(* IEC 61131-3 sources: plc_NativeGateway/src (part 2) *)

(* ---- NG_HmiEdit.st ---- *)
FUNCTION_BLOCK NG_HmiEdit
VAR_INPUT
    Busy : BOOL;
    StoreBusy : BOOL;
    Managed : BOOL;
    LocalRevision : ULINT;
    NowMs : ULINT;
END_VAR
VAR_IN_OUT
    Hmi : NG_Hmi;
    Active : NG_Config;
    Bootstrap : NG_Bootstrap;
    States : ARRAY[1..50] OF NG_MeterState;
    Samples : ARRAY[1..320] OF NG_Sample;
END_VAR
VAR_OUTPUT
    Submit : BOOL;
    SubmitBroker : BOOL;
    SubmitMode : BOOL;
    SubmitReset : BOOL;
    ClearConfig : BOOL;
    Draft : NG_Config;
    NewBroker : NG_Bootstrap;
    NewManaged : BOOL;
END_VAR
VAR
    Change : NG_EditDevice;
    EditPoints : ARRAY[1..32] OF NG_Point;
    BlankPoint : NG_Point;
    BlankDevice : NG_Device;
    BaseVersion : ULINT;
    BaseRevision : ULINT;
    ModeTargetManaged : BOOL;
    ModeReviewOpen : BOOL;
    ResetReviewOpen : BOOL;
    Initialized : BOOL;
    Dirty : BOOL;
    Awaiting : BOOL;
    Reload : BOOL;
    LoadDevice : BOOL;
    LoadPoint : BOOL;
    ValidBroker : BOOL;
    RefreshAt : ULINT;
    Nav : STRING[16];
    d : INT;
    p : INT;
    i : INT;
    row : INT;
    a : INT;
    b : INT;
    idx : INT;
    pages : INT;
    point : NG_Point;
    device : NG_Device;
    rows : ARRAY[1..8] OF NG_UiLabel;
    marker : STRING[3];
    status : STRING[24];
    value : STRING[64];
    cmd : BOOL;
    Utf8 : NG_Utf8Label;
    DeviceLabel : NG_UiLabel;
    PointLabel : NG_UiLabel;
    UnitLabel : NG_UiLabel;
END_VAR
Submit := FALSE; SubmitBroker := FALSE; SubmitMode := FALSE; SubmitReset := FALSE; ClearConfig := FALSE; LoadDevice := FALSE; LoadPoint := FALSE;
Nav := Hmi.Navigation; Hmi.Navigation := '';
IF Nav='ZH' THEN Hmi.English:=FALSE;
ELSIF Nav='EN' THEN Hmi.English:=TRUE;
ELSIF Nav='REFRESH' THEN IF Dirty THEN Hmi.View:=5; ELSE Hmi.Load:=TRUE; END_IF;
ELSIF Nav='DISCARD' THEN Hmi.Load:=TRUE; Hmi.View:=0;
ELSIF Nav='REVIEW' THEN Hmi.View:=6;
ELSIF Nav='COMMIT' THEN Hmi.Apply:=TRUE;
ELSIF Nav='DEVON' THEN Hmi.DeviceEnabled:='true';
ELSIF Nav='DEVOFF' THEN Hmi.DeviceEnabled:='false';
ELSIF Nav='POINTON' THEN Hmi.PointEnabled:='true';
ELSIF Nav='POINTOFF' THEN Hmi.PointEnabled:='false';
ELSIF Nav='MODEPAGE' THEN ModeReviewOpen:=FALSE; ResetReviewOpen:=FALSE; Hmi.View:=13;
ELSIF Nav='MODEHUB' THEN ModeTargetManaged:=TRUE; ModeReviewOpen:=TRUE; ResetReviewOpen:=FALSE; Hmi.ClearOnMaintenance:=FALSE; Hmi.View:=15;
ELSIF Nav='MODELOCAL' THEN ModeTargetManaged:=FALSE; ModeReviewOpen:=TRUE; ResetReviewOpen:=FALSE; Hmi.ClearOnMaintenance:=FALSE; Hmi.View:=14;
ELSIF Nav='MODEKEEP' THEN Hmi.ClearOnMaintenance:=FALSE;
ELSIF Nav='MODECLEAR' THEN Hmi.ClearOnMaintenance:=TRUE;
ELSIF Nav='MODECOMMIT' THEN
    IF ModeReviewOpen AND ((Hmi.View=14) OR (Hmi.View=15)) THEN Hmi.SwitchMode:=TRUE;
    ELSE Hmi.Status:='Open the management mode confirmation before saving.'; END_IF;
ELSIF Nav='RESETPAGE' THEN ModeReviewOpen:=FALSE; ResetReviewOpen:=TRUE; Hmi.View:=16;
ELSIF Nav='RESETCOMMIT' THEN
    IF ResetReviewOpen AND (Hmi.View=16) THEN
        IF StoreBusy THEN Hmi.Status:='Busy: configuration transaction in progress. Try again shortly.';
        ELSE SubmitReset:=TRUE; ResetReviewOpen:=FALSE; Dirty:=FALSE; Awaiting:=FALSE; Reload:=TRUE; Hmi.View:=0; Hmi.Status:='Clearing local configuration and version baseline...'; END_IF;
    ELSE Hmi.Status:='Open the reset confirmation before clearing local configuration.'; END_IF;
ELSIF Nav='CYCLIC' THEN Hmi.ReportMode:='cyclic';
ELSIF Nav='CHANGE' THEN Hmi.ReportMode:='change';
ELSIF Nav='BOTH' THEN Hmi.ReportMode:='change_or_cyclic';
ELSIF Nav='HOLDING' THEN Hmi.Area:='holding_register';
ELSIF Nav='INPUT' THEN Hmi.Area:='input_register';
ELSIF Nav='COIL' THEN Hmi.Area:='coil';
ELSIF Nav='DISCRETE' THEN Hmi.Area:='discrete_input';
ELSIF Nav='UINT16' THEN Hmi.DataType:='uint16'; Hmi.ByteOrder:='AB';
ELSIF Nav='INT16' THEN Hmi.DataType:='int16'; Hmi.ByteOrder:='AB';
ELSIF Nav='UINT32' THEN Hmi.DataType:='uint32'; Hmi.ByteOrder:='ABCD';
ELSIF Nav='INT32' THEN Hmi.DataType:='int32'; Hmi.ByteOrder:='ABCD';
ELSIF Nav='FLOAT32' THEN Hmi.DataType:='float32'; Hmi.ByteOrder:='ABCD';
ELSIF Nav='BOOL' THEN Hmi.DataType:='bool'; Hmi.ByteOrder:=''; Hmi.Scale:='1'; Hmi.Offset:='0'; Hmi.Deadband:='0';
ELSIF Nav='ADVANCED' THEN Hmi.Advanced:=NOT Hmi.Advanced;
ELSIF Nav='BROKERREVIEW' THEN Hmi.View:=7;
ELSIF Nav='BROKERCOMMIT' THEN Hmi.SaveBroker:=TRUE;
ELSIF Nav='HELP' THEN Hmi.View:=8;
ELSIF Nav='TYPEPICK' THEN Hmi.View:=9;
ELSIF Nav='AREAPICK' THEN Hmi.View:=10;
ELSIF Nav='REPORTPICK' THEN Hmi.View:=11;
ELSIF Nav='GATEWAY' THEN Hmi.View:=12;
ELSIF Nav='POINTBACK' THEN Hmi.View:=2;
END_IF;
IF (Nav='CYCLIC') OR (Nav='CHANGE') OR (Nav='BOTH') OR (Nav='HOLDING') OR (Nav='INPUT') OR (Nav='COIL') OR (Nav='DISCRETE') OR (Nav='UINT16') OR (Nav='INT16') OR (Nav='UINT32') OR (Nav='INT32') OR (Nav='FLOAT32') OR (Nav='BOOL') THEN Hmi.View:=2; END_IF;
Hmi.Managed:=Managed;
IF Managed THEN Hmi.ManagementMode:='HUB_MANAGED'; ELSE Hmi.ManagementMode:='STANDALONE'; END_IF;
IF Managed AND ((Nav='DNEW') OR (Nav='PNEW') OR (Nav='DDEL') OR (Nav='PDEL') OR (Nav='PERIOD') OR Hmi.SaveDevice OR Hmi.SavePoint OR Hmi.RemoveDevice OR Hmi.RemovePoint OR Hmi.Apply) THEN
    Nav := ''; Hmi.SaveDevice:=FALSE; Hmi.SavePoint:=FALSE; Hmi.RemoveDevice:=FALSE; Hmi.RemovePoint:=FALSE; Hmi.Apply:=FALSE;
    Hmi.View:=0; Hmi.Status:='HUB_MANAGED: publish device and point changes from Hub.';
END_IF;
IF Managed THEN Hmi.ConfigSource:='HUB_MANAGED - local device/point changes blocked'; ELSE Hmi.ConfigSource:='MAINTENANCE - incoming platform configuration locked'; END_IF;
IF NOT Initialized THEN Reload := TRUE; Initialized := TRUE; END_IF;
IF Awaiting AND (Active.Version = Draft.Version) AND NOT Busy THEN Dirty := FALSE; Awaiting := FALSE; Reload := TRUE; Hmi.View:=0; END_IF;
IF ((Active.Version <> BaseVersion) OR (LocalRevision <> BaseRevision)) AND NOT Dirty AND NOT Awaiting AND NOT Busy THEN Reload := TRUE; END_IF;
IF Hmi.Load AND NOT Busy THEN Reload := TRUE; Hmi.View:=0; Hmi.Status := 'Display refreshed from active configuration. Unapplied draft discarded.'; END_IF;
IF Reload THEN
    Draft := Active; BaseVersion := Active.Version; BaseRevision := LocalRevision; Dirty := FALSE; Reload := FALSE;
    Hmi.Enabled := TO_STRING(Draft.enabled,''); Hmi.BatchIntervalMs := TO_STRING(Draft.batchIntervalMs,'{0:d}'); Hmi.MaxBatchPoints := TO_STRING(Draft.maxBatchPoints,'{0:d}');
    IF NOT NG_Range(Hmi.DeviceIndex,1,50,TRUE) THEN Hmi.DeviceIndex := '1'; END_IF;
    Hmi.PointIndex := '1'; LoadDevice := TRUE; LoadPoint := TRUE;
END_IF;
d := 1; p := 1;
IF NG_Range(Hmi.DeviceIndex,1,50,TRUE) THEN d := TO_INT(Hmi.DeviceIndex); END_IF;
IF NG_Range(Hmi.PointIndex,1,32,TRUE) THEN p := TO_INT(Hmi.PointIndex); END_IF;
IF Nav = 'LIST' THEN Hmi.View := 0;
ELSIF Nav = 'MQTT' THEN Hmi.View := 3;
ELSIF Nav = 'DEDIT' THEN Hmi.View := 1; LoadDevice := TRUE;
ELSIF Nav = 'PEDIT' THEN Hmi.View := 2; LoadPoint := TRUE;
ELSIF Nav = 'DPREV' THEN Hmi.DevicePage := MAX(1,Hmi.DevicePage-1);
ELSIF Nav = 'DNEXT' THEN Hmi.DevicePage := MIN(MAX(1,(Draft.DeviceCount+7)/8),Hmi.DevicePage+1);
ELSIF Nav = 'PPREV' THEN Hmi.PointPage := MAX(1,Hmi.PointPage-1);
ELSIF Nav = 'PNEXT' THEN IF d <= Draft.DeviceCount THEN Hmi.PointPage := MIN(MAX(1,(Draft.Devices[d].PointCount+7)/8),Hmi.PointPage+1); END_IF;
ELSIF Nav = 'DDEL' THEN Hmi.DeleteKind := 1; Hmi.View := 4;
ELSIF Nav = 'PDEL' THEN Hmi.DeleteKind := 2; Hmi.View := 4;
ELSIF Nav = 'CANCEL' THEN Hmi.DeleteKind := 0; Hmi.View := 0;
ELSIF Nav = 'DNEW' THEN
    IF Draft.DeviceCount >= 50 THEN Hmi.Status := 'Capacity reached: 50 devices.';
    ELSE
        d := Draft.DeviceCount+1; Hmi.DeviceIndex := TO_STRING(d,'{0:d}'); Hmi.PointIndex := '1'; Hmi.View := 1;
        Hmi.DeviceId := CONCAT('meter-',TO_STRING(d,'{0:d}')); Hmi.DeviceName := CONCAT('Meter ',TO_STRING(d,'{0:d}'));
        Hmi.Host := '192.168.0.5'; Hmi.Port := '11502'; Hmi.UnitId := TO_STRING(d,'{0:d}'); Hmi.DeviceEnabled := 'true';
        Hmi.ConnectTimeoutMs := '3000'; Hmi.RequestTimeoutMs := '1500'; Hmi.RetryCount := '0';
        Hmi.Status := 'New device: save into draft, then add its points.';
    END_IF;
ELSIF Nav = 'PNEW' THEN
    IF d > Draft.DeviceCount THEN Hmi.Status := 'Save a device into the draft first.';
    ELSIF (Draft.Devices[d].PointCount >= 32) OR (Draft.PointCount >= 320) THEN Hmi.Status := 'Capacity reached: 32 points/device, 320 shared points.';
    ELSE
        p := Draft.Devices[d].PointCount+1; Hmi.PointIndex := TO_STRING(p,'{0:d}'); Hmi.View := 2;
        Hmi.PointId := CONCAT('point-',TO_STRING(p,'{0:d}')); Hmi.PointName := CONCAT('Point ',TO_STRING(p,'{0:d}')); Hmi.PointEnabled := 'true';
        Hmi.DataType := 'float32'; Hmi.Area := 'input_register'; Hmi.Address := TO_STRING((p-1)*2,'{0:d}'); Hmi.ByteOrder := 'ABCD';
        Hmi.PollIntervalMs := '5000'; Hmi.ReportIntervalMs := '5000'; Hmi.Scale := '1'; Hmi.Offset := '0'; Hmi.Unit := '';
        Hmi.ReportMode := 'cyclic'; Hmi.Deadband := '0'; Hmi.StaleAfterMs := '20000';
        Hmi.Status := 'New point: save into draft, then apply the complete draft.';
    END_IF;
ELSIF LEN(Nav) = 2 THEN
    IF (LEFT(Nav,1) = 'D') AND NG_Range(RIGHT(Nav,1),1,8,TRUE) THEN
        i := (Hmi.DevicePage-1)*8+TO_INT(RIGHT(Nav,1));
        IF i <= Draft.DeviceCount THEN d := i; p := 1; Hmi.DeviceIndex := TO_STRING(d,'{0:d}'); Hmi.PointIndex := '1'; Hmi.PointPage := 1; LoadDevice := TRUE; LoadPoint := TRUE; END_IF;
    ELSIF (LEFT(Nav,1) = 'P') AND NG_Range(RIGHT(Nav,1),1,8,TRUE) AND (d <= Draft.DeviceCount) THEN
        i := (Hmi.PointPage-1)*8+TO_INT(RIGHT(Nav,1));
        IF i <= Draft.Devices[d].PointCount THEN p := i; Hmi.PointIndex := TO_STRING(p,'{0:d}'); LoadPoint := TRUE; END_IF;
    END_IF;
END_IF;
IF LoadDevice AND (d <= Draft.DeviceCount) THEN
    device := Draft.Devices[d];
    Hmi.DeviceId := device.deviceId; Hmi.DeviceName := device.name; Hmi.DeviceEnabled := TO_STRING(device.enabled,''); Hmi.Host := device.host;
    Hmi.Port := TO_STRING(device.port,'{0:d}'); Hmi.UnitId := TO_STRING(device.unitId,'{0:d}'); Hmi.ConnectTimeoutMs := TO_STRING(device.connectTimeoutMs,'{0:d}');
    Hmi.RequestTimeoutMs := TO_STRING(device.requestTimeoutMs,'{0:d}'); Hmi.RetryCount := TO_STRING(device.retryCount,'{0:d}');
END_IF;
IF Hmi.LoadPoint THEN LoadPoint := TRUE; END_IF;
IF LoadPoint AND (d <= Draft.DeviceCount) THEN
    IF p <= Draft.Devices[d].PointCount THEN
        point := Draft.Points[Draft.Devices[d].PointStart+p-1];
        Hmi.PointId := point.pointId; Hmi.PointName := point.name; Hmi.PointEnabled := TO_STRING(point.enabled,''); Hmi.DataType := point.dataType;
        Hmi.PollIntervalMs := TO_STRING(point.pollIntervalMs,'{0:d}'); Hmi.ReportIntervalMs := TO_STRING(point.reportIntervalMs,'{0:d}');
        Hmi.Scale := TO_STRING(point.scale,'{0:F6}'); Hmi.Offset := TO_STRING(point.offset,'{0:F6}'); Hmi.Unit := point.unit; Hmi.ReportMode := point.reportMode;
        Hmi.Deadband := TO_STRING(point.deadband,'{0:F6}'); Hmi.StaleAfterMs := TO_STRING(point.staleAfterMs,'{0:d}'); Hmi.Area := point.area;
        Hmi.Address := TO_STRING(point.address,'{0:d}'); Hmi.ByteOrder := point.byteOrder;
        Hmi.DevicePollMs := Hmi.PollIntervalMs; Hmi.DeviceReportMs := Hmi.ReportIntervalMs;
    END_IF;
END_IF;
cmd := Hmi.SaveDevice OR Hmi.SavePoint OR Hmi.RemoveDevice OR Hmi.RemovePoint OR Hmi.Apply OR Hmi.SaveBroker OR Hmi.SwitchMode OR (Nav = 'PERIOD');
IF cmd AND ((Hmi.SaveBroker AND StoreBusy) OR ((NOT Hmi.SaveBroker) AND Busy)) THEN Hmi.Status := 'Busy: configuration transaction in progress. Try again shortly.';
ELSIF cmd THEN
    IF NOT NG_Range(Hmi.DeviceIndex,1,50,TRUE) OR NOT NG_Range(Hmi.PointIndex,1,32,TRUE) THEN Hmi.Status := 'Device index 1..50; point index 1..32.';
    ELSE
        d := TO_INT(Hmi.DeviceIndex); p := TO_INT(Hmi.PointIndex); device := BlankDevice;
        IF d <= Draft.DeviceCount THEN device := Draft.Devices[d]; FOR i := 1 TO device.PointCount DO EditPoints[i] := Draft.Points[device.PointStart+i-1]; END_FOR; END_IF;
        IF Hmi.SaveDevice THEN
            IF (d > Draft.DeviceCount+1) OR NOT NG_ValidId(Hmi.DeviceId) OR (LEN(Hmi.DeviceName)=0) OR NOT NG_IPv4(Hmi.Host) OR
               NOT NG_Range(Hmi.Port,1,65535,TRUE) OR NOT NG_Range(Hmi.UnitId,0,255,TRUE) OR NOT NG_Range(Hmi.ConnectTimeoutMs,1,300000,TRUE) OR NOT NG_Range(Hmi.RequestTimeoutMs,1,300000,TRUE) OR NOT NG_Range(Hmi.RetryCount,0,10,TRUE) THEN Hmi.Status := 'Invalid device fields: check ID, name, IPv4, port and timeout values.';
            ELSE
                device.deviceId := Hmi.DeviceId; device.name := Hmi.DeviceName; device.enabled := (Hmi.DeviceEnabled='true') OR (Hmi.DeviceEnabled='TRUE');
                device.host := Hmi.Host; device.port := TO_UINT(Hmi.Port); device.unitId := TO_USINT(Hmi.UnitId); device.connectTimeoutMs := TO_UDINT(Hmi.ConnectTimeoutMs);
                device.requestTimeoutMs := TO_UDINT(Hmi.RequestTimeoutMs); device.retryCount := TO_USINT(Hmi.RetryCount);
                Change(DeviceIndex := d, Remove := FALSE, Replacement := device, Config := Draft, Points := EditPoints);
                IF Change.ErrorText = '' THEN Dirty := TRUE; Hmi.View := 0; Hmi.Status := 'Device saved to draft. Apply draft to persist.'; ELSE Hmi.Status := Change.ErrorText; END_IF;
            END_IF;
        END_IF;
        IF Hmi.SavePoint THEN
            IF (d > Draft.DeviceCount) OR (p > device.PointCount+1) OR NOT NG_ValidId(Hmi.PointId) OR (LEN(Hmi.PointName)=0) OR
               NOT NG_Range(Hmi.PollIntervalMs,1,86400000,TRUE) OR NOT NG_Range(Hmi.ReportIntervalMs,1,86400000,TRUE) OR NOT NG_Range(Hmi.StaleAfterMs,1,86400000,TRUE) OR NOT NG_Range(Hmi.Address,0,65535,TRUE) OR
               NOT NG_Range(Hmi.Scale,-1.0E20,1.0E20,FALSE) OR NOT NG_Range(Hmi.Offset,-1.0E20,1.0E20,FALSE) OR NOT NG_Range(Hmi.Deadband,0,1.0E20,FALSE) THEN Hmi.Status := 'Invalid point fields; save the device first and check numeric fields.';
            ELSE
                point := BlankPoint; point.pointId := Hmi.PointId; point.name := Hmi.PointName; point.enabled := (Hmi.PointEnabled='true') OR (Hmi.PointEnabled='TRUE');
                point.dataType := Hmi.DataType; point.pollIntervalMs := TO_UDINT(Hmi.PollIntervalMs); point.reportIntervalMs := TO_UDINT(Hmi.ReportIntervalMs);
                point.scale := TO_LREAL(Hmi.Scale); point.offset := TO_LREAL(Hmi.Offset); point.unit := Hmi.Unit; point.reportMode := Hmi.ReportMode;
                point.deadband := TO_LREAL(Hmi.Deadband); point.staleAfterMs := TO_UDINT(Hmi.StaleAfterMs); point.area := Hmi.Area; point.address := TO_UINT(Hmi.Address); point.byteOrder := Hmi.ByteOrder;
                EditPoints[p] := point; IF p > device.PointCount THEN device.PointCount := p; END_IF;
                Change(DeviceIndex := d, Remove := FALSE, Replacement := device, Config := Draft, Points := EditPoints);
                IF Change.ErrorText = '' THEN Dirty := TRUE; Hmi.View := 0; Hmi.Status := 'Point saved to draft. Apply draft to persist.'; ELSE Hmi.Status := Change.ErrorText; END_IF;
            END_IF;
        END_IF;
        IF Hmi.RemoveDevice AND (d <= Draft.DeviceCount) THEN
            Change(DeviceIndex := d, Remove := TRUE, Replacement := device, Config := Draft, Points := EditPoints);
            IF Change.ErrorText = '' THEN Dirty := TRUE; Hmi.DeviceIndex := '1'; Hmi.PointIndex := '1'; Hmi.View := 0; Hmi.DeleteKind := 0; Hmi.Status := 'Device and points removed from draft. Apply to persist.'; END_IF;
        END_IF;
        IF Hmi.RemovePoint AND (d <= Draft.DeviceCount) AND (p <= device.PointCount) THEN
            FOR i := p TO device.PointCount-1 DO EditPoints[i] := EditPoints[i+1]; END_FOR; device.PointCount := device.PointCount-1;
            Change(DeviceIndex := d, Remove := FALSE, Replacement := device, Config := Draft, Points := EditPoints);
            IF Change.ErrorText = '' THEN Dirty := TRUE; Hmi.PointIndex := '1'; Hmi.View := 0; Hmi.DeleteKind := 0; Hmi.Status := 'Point removed from draft. Apply to persist.'; END_IF;
        END_IF;
        IF (Nav = 'PERIOD') AND (d <= Draft.DeviceCount) THEN
            IF NOT NG_Range(Hmi.DevicePollMs,1,28800000,TRUE) OR NOT NG_Range(Hmi.DeviceReportMs,1,86400000,TRUE) THEN Hmi.Status := 'Invalid device polling/report period.';
            ELSE
                FOR i := 1 TO device.PointCount DO idx := device.PointStart+i-1; Draft.Points[idx].pollIntervalMs := TO_UDINT(Hmi.DevicePollMs); Draft.Points[idx].reportIntervalMs := TO_UDINT(Hmi.DeviceReportMs); Draft.Points[idx].staleAfterMs := MAX(Draft.Points[idx].staleAfterMs,Draft.Points[idx].pollIntervalMs*3); END_FOR;
                Dirty := TRUE; Hmi.Status := 'Device point periods updated in draft. Apply to persist.';
            END_IF;
        END_IF;
        IF Hmi.Apply THEN
            IF (BaseVersion <> Active.Version) OR (BaseRevision <> LocalRevision) THEN Hmi.Status := 'VERSION_CONFLICT: reload active configuration before applying.';
            ELSIF NOT NG_Range(Hmi.BatchIntervalMs,1,86400000,TRUE) OR NOT NG_Range(Hmi.MaxBatchPoints,1,64,TRUE) THEN Hmi.Status := 'Invalid gateway batch settings.';
            ELSE
                Draft.enabled := (Hmi.Enabled='true') OR (Hmi.Enabled='TRUE'); Draft.batchIntervalMs := TO_UDINT(Hmi.BatchIntervalMs); Draft.maxBatchPoints := TO_UINT(Hmi.MaxBatchPoints); Hmi.Status := NG_CheckConfig(Draft);
                IF Hmi.Status = '' THEN Draft.Version := Active.Version; Submit := TRUE; Awaiting := TRUE; Dirty := TRUE; Hmi.Status := 'Saving, hashing and reading back configuration...'; END_IF;
            END_IF;
        END_IF;
        IF Hmi.SwitchMode THEN
            NewManaged := ModeTargetManaged;
            IF NewManaged = Managed THEN Hmi.Status := 'The selected management mode is already active.';
            ELSE
                ClearConfig := NOT NewManaged AND Hmi.ClearOnMaintenance;
                SubmitMode := TRUE; ModeReviewOpen:=FALSE; Dirty := FALSE; Awaiting := FALSE; Reload := TRUE;
                Hmi.View := 13; Hmi.Status := 'Saving management mode; existing identity is retained.';
            END_IF;
        END_IF;
        IF Hmi.SaveBroker THEN
            ValidBroker := FALSE;
            IF LEN(Hmi.BrokerUri) >= 6 THEN ValidBroker := (LEFT(Hmi.BrokerUri,6)='tcp://') OR (LEFT(Hmi.BrokerUri,6)='ssl://'); END_IF;
            IF NOT ValidBroker OR NOT NG_ValidId(Hmi.BrokerGatewayId) OR ((Hmi.ManagementMode<>'HUB_MANAGED') AND (Hmi.ManagementMode<>'STANDALONE')) OR NOT NG_Range(Hmi.UtcOffsetMinutes,-840,840,TRUE) THEN Hmi.Status := 'Check broker URI, gateway ID, client ID and time zone.';
            ELSE
                NewManaged := Managed; NewBroker := Bootstrap; NewBroker.GatewayId:=Hmi.BrokerGatewayId; NewBroker.BrokerUri := Hmi.BrokerUri; NewBroker.ClientId := Hmi.BrokerGatewayId; Hmi.ClientId := Hmi.BrokerGatewayId; NewBroker.UserName := Hmi.UserName; NewBroker.UtcOffsetMinutes := TO_INT(Hmi.UtcOffsetMinutes);
                IF Hmi.Password <> '' THEN NewBroker.Password := Hmi.Password; END_IF;
                SubmitBroker := TRUE; Hmi.Password := ''; Hmi.View:=3; Hmi.Status := 'Saving broker settings...';
            END_IF;
        END_IF;
    END_IF;
END_IF;
Hmi.Load := FALSE; Hmi.LoadPoint := FALSE; Hmi.SaveDevice := FALSE; Hmi.SavePoint := FALSE; Hmi.RemoveDevice := FALSE; Hmi.RemovePoint := FALSE; Hmi.Apply := FALSE; Hmi.SaveBroker := FALSE; Hmi.SwitchMode := FALSE;
Hmi.UiStatus:=NG_UiText(Hmi.Status,Hmi.English);
Hmi.UiDeviceEnabled:=NG_UiText(Hmi.DeviceEnabled,Hmi.English); Hmi.UiPointEnabled:=NG_UiText(Hmi.PointEnabled,Hmi.English);
Hmi.UiArea:=NG_UiText(Hmi.Area,Hmi.English); Hmi.UiReportMode:=NG_UiText(Hmi.ReportMode,Hmi.English); Hmi.UiManagementMode:=NG_UiText(Hmi.ManagementMode,Hmi.English);
IF Dirty THEN Hmi.DraftState := 'UNSAVED DRAFT'; ELSE Hmi.DraftState := 'PERSISTED'; END_IF;
IF Dirty AND ((BaseVersion <> Active.Version) OR (BaseRevision <> LocalRevision)) AND NOT Awaiting THEN Hmi.DraftState := 'VERSION CONFLICT'; END_IF;
Hmi.UiDraftState:=NG_UiText(Hmi.DraftState,Hmi.English);
Hmi.UiConfigSource:=NG_UiText(Hmi.ConfigSource,Hmi.English);
Hmi.TotalPoints := TO_STRING(Active.PointCount,'{0:d}');
IF (NowMs < RefreshAt) AND (Nav = '') AND NOT cmd THEN RETURN; END_IF;
RefreshAt := NowMs+250;
Hmi.DevicePage := MAX(1,MIN(MAX(1,(Draft.DeviceCount+7)/8),Hmi.DevicePage));
Hmi.DevicePages := CONCAT(TO_STRING(Hmi.DevicePage,'{0:d}'),' / ',TO_STRING(MAX(1,(Draft.DeviceCount+7)/8),'{0:d}'));
FOR row := 1 TO 8 DO
    i := (Hmi.DevicePage-1)*8+row; rows[row] := "";
    IF i <= Draft.DeviceCount THEN
        device := Draft.Devices[i]; marker := ''; IF i = d THEN marker := '> '; END_IF;
        status := 'DRAFT'; FOR a := 1 TO Active.DeviceCount DO IF Active.Devices[a].deviceId = device.deviceId THEN status := States[a].StateText; EXIT; END_IF; END_FOR;
        Utf8(Text := device.name, MaxChars := 48); DeviceLabel := Utf8.Value;
        IF Hmi.English THEN
            rows[row]:=NG_UiJoin(TO_WSTRING(marker,""),DeviceLabel," | ",NG_UiText(status,TRUE),"\n",TO_WSTRING(CONCAT(device.host,':',TO_STRING(device.port,'{0:d}')),""),TO_WSTRING(device.unitId," / Unit {0:d}"),TO_WSTRING(device.PointCount," / {0:d} points"));
        ELSE
            rows[row]:=NG_UiJoin(TO_WSTRING(marker,""),DeviceLabel," | ",NG_UiText(status,FALSE),"\n",TO_WSTRING(CONCAT(device.host,':',TO_STRING(device.port,'{0:d}')),""),TO_WSTRING(device.unitId," / 站号 {0:d}"),TO_WSTRING(device.PointCount," / {0:d} 个点位"));
        END_IF;
    END_IF;
END_FOR;
Hmi.DeviceRow1 := rows[1]; Hmi.DeviceRow2 := rows[2]; Hmi.DeviceRow3 := rows[3]; Hmi.DeviceRow4 := rows[4]; Hmi.DeviceRow5 := rows[5]; Hmi.DeviceRow6 := rows[6]; Hmi.DeviceRow7 := rows[7]; Hmi.DeviceRow8 := rows[8];
Hmi.SelectedDevice := NG_UiText('No device selected',Hmi.English); Hmi.SelectedPoint := NG_UiText('No point selected',Hmi.English);
IF d <= Draft.DeviceCount THEN Utf8(Text := Draft.Devices[d].name, MaxChars := 0); Hmi.SelectedDevice := Utf8.Value; END_IF;
pages := 1; IF d <= Draft.DeviceCount THEN pages := MAX(1,(Draft.Devices[d].PointCount+7)/8); END_IF;
Hmi.PointPage := MAX(1,MIN(pages,Hmi.PointPage)); Hmi.PointPages := CONCAT(TO_STRING(Hmi.PointPage,'{0:d}'),' / ',TO_STRING(pages,'{0:d}'));
FOR row := 1 TO 8 DO
    i := (Hmi.PointPage-1)*8+row; rows[row] := "";
    IF d <= Draft.DeviceCount THEN
        IF i <= Draft.Devices[d].PointCount THEN
            point := Draft.Points[Draft.Devices[d].PointStart+i-1]; marker := '';
            IF (point.name='voltage') OR (point.name='current') OR (point.name='frequency') OR (point.name='power') OR (point.name='energy') THEN
                PointLabel := NG_UiText(point.name,Hmi.English);
            ELSE
                Utf8(Text := point.name, MaxChars := 0); PointLabel := Utf8.Value;
            END_IF;
            IF i = p THEN marker := '> '; Hmi.SelectedPoint := PointLabel; END_IF;
            status := 'DRAFT'; value := '';
            FOR a := 1 TO Active.DeviceCount DO
                IF Active.Devices[a].deviceId = Draft.Devices[d].deviceId THEN
                    FOR b := 1 TO Active.Devices[a].PointCount DO idx := Active.Devices[a].PointStart+b-1; IF Active.Points[idx].pointId = point.pointId THEN status := Samples[idx].Quality; IF status = 'GOOD' THEN IF ABS(Samples[idx].Value)<1.0E9 THEN value := TO_STRING(Samples[idx].Value,'{0:F3}'); ELSE value := TO_STRING(Samples[idx].Value,'{0:E6}'); END_IF; END_IF; EXIT; END_IF; END_FOR; EXIT;
                END_IF;
            END_FOR;
            Utf8(Text := CONCAT(value,' ',point.unit), MaxChars := 0); UnitLabel := Utf8.Value;
            rows[row]:=NG_UiJoin(TO_WSTRING(marker,""),PointLabel,"  |  ",UnitLabel,"  |  ",NG_UiText(status,Hmi.English),"\n",NG_UiText(point.area,Hmi.English));
            IF Hmi.English THEN
                rows[row]:=NG_UiJoin(rows[row],TO_WSTRING(point.address," @{0:d}"),TO_WSTRING(point.pollIntervalMs," / Poll {0:d}"),TO_WSTRING(point.reportIntervalMs," / Send {0:d} ms"),"","","","");
            ELSE
                rows[row]:=NG_UiJoin(rows[row],TO_WSTRING(point.address," @{0:d}"),TO_WSTRING(point.pollIntervalMs," / 采集 {0:d}"),TO_WSTRING(point.reportIntervalMs," / 上报 {0:d} 毫秒"),"","","","");
            END_IF;
        END_IF;
    END_IF;
END_FOR;
Hmi.PointRow1 := rows[1]; Hmi.PointRow2 := rows[2]; Hmi.PointRow3 := rows[3]; Hmi.PointRow4 := rows[4]; Hmi.PointRow5 := rows[5]; Hmi.PointRow6 := rows[6]; Hmi.PointRow7 := rows[7]; Hmi.PointRow8 := rows[8];
END_FUNCTION_BLOCK

(* ---- NG_JsonParse.st ---- *)
FUNCTION_BLOCK NG_JsonParse
VAR_INPUT
    Execute : BOOL;
    Length : UDINT;
END_VAR
VAR_IN_OUT
    Buffer : NG_Bytes;
    Doc : NG_Document;
END_VAR
VAR_OUTPUT
    Done : BOOL;
    Busy : BOOL;
    Error : BOOL;
    ErrorText : NG_Text;
END_VAR
VAR
    ConvertChar : NG_Char;
    Previous : BOOL;
    Pos : DINT;
    Depth : INT;
    Nodes : ARRAY[0..64] OF INT;
    Expected : ARRAY[0..64] OF INT;
    Keys : ARRAY[0..64] OF NG_Id;
    Mode : INT;
    IsKey : BOOL;
    Text : STRING[512];
    Start : DINT;
    Code : UINT;
    UCode : UDINT;
    HighSurrogate : UDINT;
    HexCount : INT;
    N : INT;
    I : INT;
    Budget : INT;
    C : STRING[1];
    Again : BOOL;
    FinishScalar : BOOL;
    Kind : INT;
    NewValue : BOOL;
    Parent : INT;
    Number : LREAL;
    ClipIndex : INT;
END_VAR
IF Execute AND NOT Previous AND NOT Busy THEN
    Pos := 0; Depth := 0; Doc.Count := 0; Mode := 0;
    Nodes[0] := 0; Expected[0] := 2; Keys[0] := '';
    Done := FALSE; Error := FALSE; ErrorText := ''; Busy := TRUE;
    IF (Length = 0) OR (Length > 131071) THEN
        Error := TRUE; ErrorText := 'PAYLOAD_TOO_LARGE';
    END_IF;
END_IF;
Previous := Execute;
IF NOT Busy THEN RETURN; END_IF;
Budget := 0;
WHILE (Budget < 512) AND NOT Error DO
    IF Pos >= TO_DINT(Length) THEN
        IF Mode = 4 THEN FinishScalar := TRUE;
        ELSIF (Mode = 0) AND (Depth = 0) AND (Doc.Count > 0) THEN
            Done := TRUE; Busy := FALSE; EXIT;
        ELSE Error := TRUE; EXIT;
        END_IF;
        Code := 0; C := '';
    ELSE Code := TO_UINT(Buffer[Pos]); ConvertChar(Code := Code, Utf8 := FALSE); C := ConvertChar.Value;
    END_IF;
    Again := FALSE; NewValue := FALSE;
    CASE Mode OF
    0:
        IF (Code = 32) OR (Code = 9) OR (Code = 10) OR (Code = 13) THEN
            Pos := Pos + 1;
        ELSIF (Code = 125) OR (Code = 93) THEN
            IF Depth = 0 THEN Error := TRUE;
            ELSIF ((Doc.Tokens[Nodes[Depth]].Kind = 1) AND (Code = 125) AND ((Expected[Depth] = 0) OR (Expected[Depth] = 3))) OR
                  ((Doc.Tokens[Nodes[Depth]].Kind = 2) AND (Code = 93) AND ((Expected[Depth] = 5) OR (Expected[Depth] = 6))) THEN
                Doc.Tokens[Nodes[Depth]].NextToken := Doc.Count + 1;
                Depth := Depth - 1; Pos := Pos + 1;
            ELSE Error := TRUE;
            END_IF;
        ELSIF (Code = 44) AND (Depth > 0) THEN
            IF Expected[Depth] = 3 THEN Expected[Depth] := 4;
            ELSIF Expected[Depth] = 6 THEN Expected[Depth] := 7;
            ELSE Error := TRUE; END_IF;
            Pos := Pos + 1;
        ELSIF (Code = 58) AND (Expected[Depth] = 1) THEN
            Expected[Depth] := 2; Pos := Pos + 1;
        ELSIF ((Expected[Depth] = 0) OR (Expected[Depth] = 4)) AND (Code = 34) THEN
            IsKey := TRUE; Text := ''; Mode := 1; Pos := Pos + 1; HighSurrogate := 0;
        ELSIF (Expected[Depth] = 2) OR (Expected[Depth] = 5) OR (Expected[Depth] = 7) THEN
            IF Depth = 0 THEN Expected[Depth] := 8;
            ELSIF Doc.Tokens[Nodes[Depth]].Kind = 1 THEN Expected[Depth] := 3;
            ELSE Expected[Depth] := 6; END_IF;
            Start := Pos; IsKey := FALSE; Text := ''; HighSurrogate := 0;
            IF Code = 34 THEN Mode := 1; Pos := Pos + 1;
            ELSIF (Code = 123) OR (Code = 91) THEN
                IF Code = 123 THEN Kind := 1; ELSE Kind := 2; END_IF;
                NewValue := TRUE; Pos := Pos + 1;
            ELSIF (Code = 45) OR ((Code >= 48) AND (Code <= 57)) OR (Code = 116) OR (Code = 102) OR (Code = 110) THEN
                Mode := 4; Again := TRUE;
            ELSE Error := TRUE; END_IF;
        ELSE Error := TRUE;
        END_IF;
    1:
        IF Code = 34 THEN
            IF HighSurrogate <> 0 THEN Error := TRUE;
            ELSIF IsKey THEN
                IF LEN(Text) > 64 THEN Error := TRUE;
                ELSE Keys[Depth] := Text; Expected[Depth] := 1; END_IF;
            ELSE Kind := 3; NewValue := TRUE; END_IF;
            Mode := 0; Pos := Pos + 1;
        ELSIF Code = 92 THEN Mode := 2; Pos := Pos + 1;
        ELSIF (Code < 32) OR (LEN(Text) >= 512) OR (HighSurrogate <> 0) THEN Error := TRUE;
        ELSE Text := CONCAT(Text,C); Pos := Pos + 1;
        END_IF;
    2:
        IF Code = 117 THEN UCode := 0; HexCount := 0; Mode := 3;
        ELSIF HighSurrogate <> 0 THEN Error := TRUE;
        ELSIF (Code = 34) OR (Code = 92) OR (Code = 47) THEN Text := CONCAT(Text,C); Mode := 1;
        ELSIF Code = 98 THEN ConvertChar(Code := 8, Utf8 := FALSE); Text := CONCAT(Text,ConvertChar.Value); Mode := 1;
        ELSIF Code = 102 THEN ConvertChar(Code := 12, Utf8 := FALSE); Text := CONCAT(Text,ConvertChar.Value); Mode := 1;
        ELSIF Code = 110 THEN ConvertChar(Code := 10, Utf8 := FALSE); Text := CONCAT(Text,ConvertChar.Value); Mode := 1;
        ELSIF Code = 114 THEN ConvertChar(Code := 13, Utf8 := FALSE); Text := CONCAT(Text,ConvertChar.Value); Mode := 1;
        ELSIF Code = 116 THEN ConvertChar(Code := 9, Utf8 := FALSE); Text := CONCAT(Text,ConvertChar.Value); Mode := 1;
        ELSE Error := TRUE;
        END_IF;
        IF LEN(Text) > 512 THEN Error := TRUE; END_IF;
        Pos := Pos + 1;
    3:
        UCode := UCode * 16;
        IF (Code >= 48) AND (Code <= 57) THEN UCode := UCode + Code - 48;
        ELSIF (Code >= 65) AND (Code <= 70) THEN UCode := UCode + Code - 55;
        ELSIF (Code >= 97) AND (Code <= 102) THEN UCode := UCode + Code - 87;
        ELSE Error := TRUE; END_IF;
        HexCount := HexCount + 1; Pos := Pos + 1;
        IF HexCount = 4 THEN
            Mode := 1;
            IF (UCode >= 16#D800) AND (UCode <= 16#DBFF) AND (HighSurrogate = 0) THEN
                HighSurrogate := UCode;
            ELSE
                IF HighSurrogate <> 0 THEN
                    IF (UCode < 16#DC00) OR (UCode > 16#DFFF) THEN Error := TRUE;
                    ELSE UCode := UDINT#65536 + (HighSurrogate - 16#D800) * 1024 + UCode - 16#DC00;
                    END_IF;
                    HighSurrogate := 0;
                ELSIF (UCode >= 16#DC00) AND (UCode <= 16#DFFF) THEN Error := TRUE;
                END_IF;
                (* IEC strings cannot contain NUL. Reject rather than truncate. *)
                IF UCode = 0 THEN Error := TRUE;
                ELSE ConvertChar(Code := UCode, Utf8 := TRUE); Text := CONCAT(Text,ConvertChar.Value);
                END_IF;
                IF LEN(Text) > 512 THEN Error := TRUE; END_IF;
            END_IF;
        END_IF;
    4:
        IF (Pos >= TO_DINT(Length)) OR (Code = 32) OR (Code = 9) OR (Code = 10) OR (Code = 13) OR (Code = 44) OR (Code = 125) OR (Code = 93) THEN
            FinishScalar := TRUE;
        ELSIF LEN(Text) >= 128 THEN Error := TRUE;
        ELSE Text := CONCAT(Text,C); Pos := Pos + 1;
        END_IF;
    END_CASE;
    IF FinishScalar THEN
        FinishScalar := FALSE; Mode := 0; NewValue := TRUE;
        IF (Text = 'true') OR (Text = 'false') THEN Kind := 5;
        ELSIF Text = 'null' THEN Kind := 6;
        ELSIF NG_NumberValid(Text) THEN
            Kind := 4;
            (* Bound conversion exponents before the runtime conversion. *)
            IF (FIND(Text,'e') > 0) OR (FIND(Text,'E') > 0) THEN
                I := FIND(Text,'e'); IF I = 0 THEN I := FIND(Text,'E'); END_IF;
                IF ABS(TO_DINT(MID(Text,LEN(Text)-I,I+1))) > 308 THEN Error := TRUE; END_IF;
            END_IF;
            IF NOT Error THEN Number := TO_LREAL(Text); END_IF;
        ELSE Error := TRUE;
        END_IF;
    END_IF;
    IF NewValue AND NOT Error THEN
        IF Doc.Count >= 8192 THEN Error := TRUE; ErrorText := 'POINT_LIMIT_EXCEEDED';
        ELSE
            Parent := Nodes[Depth];
            IF (Parent > 0) AND (Doc.Tokens[Parent].Kind = 1) THEN
                I := Parent + 1;
                WHILE I <= Doc.Count DO
                    IF Doc.Tokens[I].Key = Keys[Depth] THEN Error := TRUE; EXIT; END_IF;
                    IF Doc.Tokens[I].NextToken <= I THEN Error := TRUE; EXIT; END_IF;
                    I := Doc.Tokens[I].NextToken;
                END_WHILE;
            END_IF;
            Doc.Count := Doc.Count + 1; N := Doc.Count;
            Doc.Tokens[N].Kind := Kind;
            Doc.Tokens[N].Parent := Parent;
            Doc.Tokens[N].Key := Keys[Depth]; Keys[Depth] := '';
            Doc.Tokens[N].TextLength := LEN(Text);
            IF LEN(Text)<=256 THEN Doc.Tokens[N].Text:=Text;
            ELSE
                (* Nested IEC string builtins use an 80-byte temporary. Copy
                   this diagnostic prefix using bounded single-byte results. *)
                Doc.Tokens[N].Text:='';
                FOR ClipIndex:=1 TO 256 DO
                    Doc.Tokens[N].Text:=CONCAT(Doc.Tokens[N].Text,MID(Text,1,ClipIndex));
                END_FOR;
            END_IF;
            Doc.Tokens[N].Number := Number;
            Doc.Tokens[N].Start := Start;
            Doc.Tokens[N].Count := Pos - Start;
            Doc.Tokens[N].NextToken := N + 1;
            IF (Kind = 1) OR (Kind = 2) THEN
                IF Depth >= 64 THEN Error := TRUE;
                ELSE
                    Depth := Depth + 1; Nodes[Depth] := N; Keys[Depth] := '';
                    IF Kind = 1 THEN Expected[Depth] := 0; ELSE Expected[Depth] := 5; END_IF;
                END_IF;
            END_IF;
        END_IF;
    END_IF;
    IF NOT Again THEN Budget := Budget + 1; END_IF;
END_WHILE;
IF Error THEN
    Busy := FALSE; Done := FALSE;
    IF ErrorText = '' THEN ErrorText := 'INVALID_JSON'; END_IF;
END_IF;
END_FUNCTION_BLOCK

(* ---- NG_Modbus.st ---- *)
FUNCTION_BLOCK NG_Modbus
VAR_INPUT
    Enable : BOOL;
    Reset : BOOL;
    NowMs : ULINT;
    UnixMs : ULINT;
    MaxMergeGap : UINT := UINT#16;
    MaxGapSpan : UINT := UINT#40;
    InterFrameGapMs : UDINT := UDINT#0;
    MaxTimeoutRetries : USINT := USINT#2;
END_VAR
VAR_IN_OUT
    Device : NG_Device;
    Points : ARRAY[1..320] OF NG_Point;
    Samples : ARRAY[1..320] OF NG_Sample;
    Buffer : NG_Buffer;
END_VAR
VAR_OUTPUT
    StateText : STRING[16];
    LastError : STRING[24];
    LastGoodTimestamp : ULINT;
    Completed : UDINT;
END_VAR
VAR
    Socket : TLS_SOCKET_2;
    Send : TLS_SEND_2;
    Receive : TLS_RECEIVE_2;
    State : INT;
    Active : BOOL;
    Scan : INT;
    Selected : INT;
    i : INT;
    j : INT;
    k : INT;
    Retry : USINT;
    Deadline : ULINT;
    RetryAt : ULINT;
    BackoffLevel : USINT;
    BackoffMs : ULINT;
    Transaction : UINT;
    FunctionCode : BYTE;
    Width : UINT;
    Tx : ARRAY[0..11] OF BYTE;
    Chunk : ARRAY[0..259] OF BYTE;
    Rx : ARRAY[0..259] OF BYTE;
    RxCount : UDINT;
    FrameLength : UDINT;
    ByteCount : UINT;
    Point : NG_Point;
    Decode : ARRAY[0..3] OF BYTE;
    UIntValue : UDINT;
    IntValue : LINT;
    FloatValue : REAL;
    ToFloat : BUF_TO_REAL;
    Value : LREAL;
    OperationFailed : BOOL;
    PointDecodeFailed : BOOL;
    FailQuality : STRING[24];
    host : STRING;
    Accepted : BOOL;
    SourceResult : NG_SourceResult;
    PollSlot : NG_PollSlot;
    Index : UINT;
    SourceMarkUs : ULINT;
    NominalDueMs : ULINT;
    RequestSlot : UINT;
    RequestConfigGeneration : UDINT;
    RequestSamplingGeneration : ULINT;
    BlockIndices : ARRAY[1..64] OF UINT;
    BlockNominalDue : ARRAY[1..64] OF ULINT;
    SavedNextDue : ARRAY[1..64] OF ULINT;
    BlockCount : INT;
    BlockStartAddr : UINT;
    BlockEndAddr : UINT;
    BlockWidth : UINT;
    BlockHasHoles : BOOL;
    HoleMergeDisabled : BOOL;
    EffectiveMaxGap : UINT;
    EffectiveGapSpan : UINT;
    EffectiveContigSpan : UINT;
    SpanLimit : UINT;
    CandIndex : UINT;
    CandWidth : UINT;
    CandEnd : UINT;
    CandGap : UINT;
    CandSpan : UINT;
    BestIndex : UINT;
    BestGap : UINT;
    BestNewStart : UINT;
    BestNewEnd : UINT;
    AlreadyInBlock : BOOL;
    MergedPass : BOOL;
    RequestSentMs : ULINT;
    LastRttMs : ULINT;
    NextTxAllowedMs : ULINT;
    TimeoutInReceive : BOOL;
    StaleDrains : USINT;
    TimeoutRetryCap : USINT;
    CanRetry : BOOL;
    RemainBytes : INT;
    RawOff : INT;
    AnyGoodInBlock : BOOL;
    AnyErrorInBlock : BOOL;
    BlockLastErr : STRING[24];
END_VAR
OperationFailed := FALSE;
host := Device.host;
IF Reset OR NOT Enable OR NOT Device.enabled THEN
    IF (State>=16) AND (State<=40) THEN
        Buffer.CancelledReadsTotal:=NG_SafeAdd(Buffer.CancelledReadsTotal,ULINT#1);
        Buffer.CancellationReason:=2;
    END_IF;
    State:=90; Selected:=0; BlockCount:=0; BlockHasHoles:=FALSE; BackoffLevel:=USINT#0;
    NextTxAllowedMs:=ULINT#0; LastRttMs:=ULINT#0; TimeoutInReceive:=FALSE; StaleDrains:=USINT#0;
    IF Reset THEN HoleMergeDisabled:=FALSE; END_IF;
END_IF;
(* Limit only new socket activation work; nominal sampling grids remain fixed.
   Already-active sockets and final physical results are never budget-blocked. *)
IF (State=0) AND Enable AND Device.enabled AND (NowMs>=RetryAt) THEN
    IF Buffer.ConnectBudget=0 THEN StateText:='WAIT_CONNECT'; RETURN; END_IF;
    Buffer.ConnectBudget:=Buffer.ConnectBudget-USINT#1;
END_IF;
Socket(ACTIVATE := (State <> 90) AND Enable AND Device.enabled AND (NowMs >= RetryAt), IS_SRV := FALSE, BIND_IP := '', BIND_PORT := UINT#0, DEST_IP := host, DEST_PORT := Device.port, START_TLS := FALSE);
Send(REQ := (State = 20) OR (State = 21), HANDLE := Socket.HANDLE, DATA_CNT := UDINT#12, SEND_SECURE := FALSE, DATA := Tx);
Receive(EN_R := (State = 30) AND Socket.ACTIVE, HANDLE := Socket.HANDLE, EXP_DATA_CNT := UDINT#0, RECEIVE_SECURE := FALSE, DATA := Chunk);
ToFloat(REQ := FALSE, BUF_FORMAT := TRUE, BUF_OFFS := 0, BUF_CNT := 4, BUFFER := Decode, DST := FloatValue);
CASE State OF
0:
    StateText := 'CONNECTING'; Deadline := NowMs + Device.connectTimeoutMs; State := 10;
10:
    IF Socket.ACTIVE THEN State := 15;
    ELSIF NowMs >= Deadline THEN
        StateText := 'OFFLINE'; LastError := 'BAD_CONNECTION';
        IF BackoffLevel < USINT#5 THEN BackoffLevel := BackoffLevel + USINT#1; END_IF;
        BackoffMs := ULINT#1000;
        FOR i := 1 TO TO_INT(BackoffLevel) DO
            IF BackoffMs < ULINT#15000 THEN BackoffMs := BackoffMs * ULINT#2; ELSE BackoffMs := ULINT#30000; END_IF;
        END_FOR;
        RetryAt := NowMs + BackoffMs + TO_ULINT(Device.unitId MOD USINT#8) * ULINT#125;
        State := 90;
        (* Charge the complete final-result loop once, including dispatch and
           index work; avoid four timer calls for each individual point. *)
        SourceMarkUs:=GET_MICROSECONDS(TRUE);
        FOR i := 1 TO Device.PointCount DO
            Index:=TO_UINT(Device.PointStart+i-1);
            IF Points[Index].enabled AND (NowMs>=Buffer.Cursors[Index].NextDueMonoMs) THEN
                PollSlot(NowMs:=NowMs, PeriodMs:=Points[Index].pollIntervalMs, Cursor:=Buffer.Cursors[Index], Buffer:=Buffer);
                NominalDueMs:=PollSlot.NominalDueMs;
                SourceResult(Index:=Index, Value:=LREAL#0.0, Quality:='BAD_CONNECTION', NowMs:=NowMs, UnixMs:=UnixMs, NominalDueMs:=NominalDueMs, ConfigSlot:=Buffer.ActiveSlot, ConfigGeneration:=Buffer.Configs[Buffer.ActiveSlot].Generation, SamplingGeneration:=Buffer.SamplingGeneration, Samples:=Samples, Buffer:=Buffer);
                Accepted:=SourceResult.Accepted;
            END_IF;
        END_FOR;
        Buffer.SourceWorkUs:=Buffer.SourceWorkUs+GET_MICROSECONDS(TRUE)-SourceMarkUs;
    END_IF;
15:
    IF NOT Socket.ACTIVE THEN State := 0;
    ELSIF (NowMs >= NextTxAllowedMs) AND (Buffer.PollStartBudget>0) THEN
        Selected := 0;
        FOR i := 1 TO Device.PointCount DO
            Scan := Scan + 1; IF Scan > Device.PointCount THEN Scan := 1; END_IF;
            IF Points[Device.PointStart+Scan-1].enabled AND (NowMs >= Samples[Device.PointStart+Scan-1].NextPollMs) THEN Selected := Scan; EXIT; END_IF;
        END_FOR;
        IF Selected > 0 THEN
            Buffer.PollStartBudget:=Buffer.PollStartBudget-USINT#1;
            Index:=TO_UINT(Device.PointStart+Selected-1);
            Point:=Points[Index]; Retry:=USINT#0; StaleDrains:=USINT#0;
            Width := UINT#1;
            IF (Point.dataType = 'float32') OR (Point.dataType = 'int32') OR (Point.dataType = 'uint32') THEN Width := UINT#2; END_IF;
            BlockCount := 1;
            BlockIndices[1] := Index;
            BlockStartAddr := Point.address;
            BlockEndAddr := Point.address + Width;
            BlockHasHoles := FALSE;
            (* Register merging for holding/input registers:
               per-device maxReadRegisters (default 120, capped at 120) and maxRegisterGap
               (default MaxMergeGap), with automatic fallback on Modbus Exception. *)
            EffectiveContigSpan := UINT#120;
            IF (Device.maxReadRegisters > UINT#0) AND (Device.maxReadRegisters < EffectiveContigSpan) THEN
                EffectiveContigSpan := Device.maxReadRegisters;
            END_IF;
            IF HoleMergeDisabled THEN EffectiveMaxGap := UINT#0;
            ELSIF Device.hasMaxRegisterGap THEN
                EffectiveMaxGap := Device.maxRegisterGap;
                IF EffectiveMaxGap > UINT#118 THEN EffectiveMaxGap := UINT#118; END_IF;
            ELSE
                EffectiveMaxGap := MaxMergeGap;
                IF EffectiveMaxGap > UINT#118 THEN EffectiveMaxGap := UINT#118; END_IF;
            END_IF;
            EffectiveGapSpan := MaxGapSpan;
            IF EffectiveGapSpan > EffectiveContigSpan THEN EffectiveGapSpan := EffectiveContigSpan; END_IF;
            IF EffectiveGapSpan < UINT#1 THEN EffectiveGapSpan := UINT#1; END_IF;
            IF ((Point.area = 'holding_register') OR (Point.area = 'input_register')) AND (Point.dataType <> 'bool') THEN
                MergedPass := TRUE;
                WHILE MergedPass AND (BlockCount < 64) DO
                    MergedPass := FALSE;
                    BestIndex := UINT#0;
                    BestGap := UINT#65535;
                    BestNewStart := BlockStartAddr;
                    BestNewEnd := BlockEndAddr;
                    FOR i := 1 TO Device.PointCount DO
                        CandIndex := TO_UINT(Device.PointStart + i - 1);
                        IF Points[CandIndex].enabled
                            AND (NowMs >= Samples[CandIndex].NextPollMs)
                            AND (Points[CandIndex].area = Point.area)
                            AND (Points[CandIndex].dataType <> 'bool')
                            AND (Points[CandIndex].pollIntervalMs = Point.pollIntervalMs)
                            AND (BlockCount < 64) THEN
                            AlreadyInBlock := FALSE;
                            FOR j := 1 TO BlockCount DO
                                IF BlockIndices[j] = CandIndex THEN AlreadyInBlock := TRUE; EXIT; END_IF;
                            END_FOR;
                            IF NOT AlreadyInBlock THEN
                                CandWidth := UINT#1;
                                IF (Points[CandIndex].dataType = 'float32') OR (Points[CandIndex].dataType = 'int32') OR (Points[CandIndex].dataType = 'uint32') THEN CandWidth := UINT#2; END_IF;
                                IF Points[CandIndex].address <= (UINT#65535 - CandWidth) THEN
                                    CandEnd := Points[CandIndex].address + CandWidth;
                                    IF Points[CandIndex].address >= BlockEndAddr THEN
                                        CandGap := Points[CandIndex].address - BlockEndAddr;
                                        CandSpan := CandEnd - BlockStartAddr;
                                        IF (NOT BlockHasHoles) AND (CandGap = UINT#0) THEN SpanLimit := EffectiveContigSpan; ELSE SpanLimit := EffectiveGapSpan; END_IF;
                                        IF (CandGap <= EffectiveMaxGap) AND (CandSpan <= SpanLimit) AND (CandGap < BestGap) THEN
                                            BestIndex := CandIndex;
                                            BestGap := CandGap;
                                            BestNewStart := BlockStartAddr;
                                            BestNewEnd := CandEnd;
                                        END_IF;
                                    ELSIF CandEnd <= BlockStartAddr THEN
                                        CandGap := BlockStartAddr - CandEnd;
                                        CandSpan := BlockEndAddr - Points[CandIndex].address;
                                        IF (NOT BlockHasHoles) AND (CandGap = UINT#0) THEN SpanLimit := EffectiveContigSpan; ELSE SpanLimit := EffectiveGapSpan; END_IF;
                                        IF (CandGap <= EffectiveMaxGap) AND (CandSpan <= SpanLimit) AND (CandGap < BestGap) THEN
                                            BestIndex := CandIndex;
                                            BestGap := CandGap;
                                            BestNewStart := Points[CandIndex].address;
                                            BestNewEnd := BlockEndAddr;
                                        END_IF;
                                    END_IF;
                                END_IF;
                            END_IF;
                        END_IF;
                    END_FOR;
                    IF BestIndex > UINT#0 THEN
                        BlockCount := BlockCount + 1;
                        BlockIndices[BlockCount] := BestIndex;
                        BlockStartAddr := BestNewStart;
                        BlockEndAddr := BestNewEnd;
                        IF BestGap > UINT#0 THEN BlockHasHoles := TRUE; END_IF;
                        MergedPass := TRUE;
                    END_IF;
                END_WHILE;
            END_IF;
            BlockWidth := BlockEndAddr - BlockStartAddr;
            SourceMarkUs:=GET_MICROSECONDS(TRUE);
            FOR k := 1 TO BlockCount DO
                CandIndex := BlockIndices[k];
                SavedNextDue[k] := Buffer.Cursors[CandIndex].NextDueMonoMs;
                PollSlot(NowMs:=NowMs, PeriodMs:=Points[CandIndex].pollIntervalMs, Cursor:=Buffer.Cursors[CandIndex], Buffer:=Buffer);
                BlockNominalDue[k] := PollSlot.NominalDueMs;
                Samples[CandIndex].NextPollMs := Buffer.Cursors[CandIndex].NextDueMonoMs;
            END_FOR;
            NominalDueMs := BlockNominalDue[1];
            Buffer.SourceWorkUs:=Buffer.SourceWorkUs+GET_MICROSECONDS(TRUE)-SourceMarkUs;
            RequestSlot:=Buffer.ActiveSlot; RequestConfigGeneration:=Buffer.Configs[RequestSlot].Generation;
            RequestSamplingGeneration:=Buffer.SamplingGeneration; State:=18;
        END_IF;
    END_IF;
16:
    IF NOT Socket.ACTIVE THEN
        OperationFailed := TRUE; FailQuality := 'BAD_CONNECTION';
    ELSIF NowMs >= NextTxAllowedMs THEN
        State := 18;
    END_IF;
18:
    Point := Points[BlockIndices[1]];
    Transaction := Transaction + 1;
    IF Point.area = 'coil' THEN FunctionCode := BYTE#1;
    ELSIF Point.area = 'discrete_input' THEN FunctionCode := BYTE#2;
    ELSIF Point.area = 'holding_register' THEN FunctionCode := BYTE#3;
    ELSE FunctionCode := BYTE#4;
    END_IF;
    Tx[0] := TO_BYTE(Transaction / 256); Tx[1] := TO_BYTE(Transaction MOD 256);
    Tx[2] := BYTE#0; Tx[3] := BYTE#0; Tx[4] := BYTE#0; Tx[5] := BYTE#6;
    Tx[6] := TO_BYTE(Device.unitId); Tx[7] := FunctionCode;
    Tx[8] := TO_BYTE(BlockStartAddr / 256); Tx[9] := TO_BYTE(BlockStartAddr MOD 256);
    Tx[10] := BYTE#0; Tx[11] := TO_BYTE(BlockWidth);
    RxCount := 0; FrameLength := 0; TimeoutInReceive := FALSE;
    RequestSentMs := NowMs;
    Deadline := NowMs + Device.requestTimeoutMs; State := 20;
20:
    IF Send.ERROR THEN OperationFailed := TRUE; FailQuality := 'BAD_CONNECTION';
    ELSIF Send.DONE THEN State := 30;
    ELSE State := 21;
    END_IF;
21:
    IF Send.ERROR THEN OperationFailed := TRUE; FailQuality := 'BAD_CONNECTION';
    ELSIF Send.DONE THEN State := 30;
    ELSIF NowMs >= Deadline THEN OperationFailed := TRUE; FailQuality := 'BAD_TIMEOUT';
    END_IF;
30:
    IF Receive.ERROR OR NOT Socket.ACTIVE THEN OperationFailed := TRUE; FailQuality := 'BAD_CONNECTION';
    ELSIF Receive.NDR THEN
        IF RxCount + Receive.DATA_CNT > 260 THEN OperationFailed := TRUE; FailQuality := 'BAD_PROTOCOL';
        ELSE
            FOR i := 0 TO TO_INT(Receive.DATA_CNT)-1 DO Rx[TO_INT(RxCount)+i] := Chunk[i]; END_FOR;
            RxCount := RxCount + Receive.DATA_CNT;
            IF RxCount >= 7 THEN
                FrameLength := UDINT#6 + TO_UDINT(Rx[4])*256 + TO_UDINT(Rx[5]);
                IF (FrameLength < 9) OR (FrameLength > 260) THEN OperationFailed := TRUE; FailQuality := 'BAD_PROTOCOL';
                ELSIF RxCount >= FrameLength THEN State := 40;
                END_IF;
            END_IF;
        END_IF;
    END_IF;
    IF (NowMs >= Deadline) AND (State = 30) THEN
        OperationFailed := TRUE; FailQuality := 'BAD_TIMEOUT'; TimeoutInReceive := TRUE;
    END_IF;
40:
    IF (RxCount >= FrameLength) AND (Rx[2] = BYTE#0) AND (Rx[3] = BYTE#0) AND (Rx[6] = Tx[6])
        AND ((Rx[0] <> Tx[0]) OR (Rx[1] <> Tx[1]))
        AND (Retry > USINT#0) AND (StaleDrains < Retry) AND (NowMs < Deadline) THEN
        (* Drain a late response frame from an earlier timed-out attempt on this socket. *)
        StaleDrains := StaleDrains + USINT#1;
        IF RxCount > FrameLength THEN
            RemainBytes := TO_INT(RxCount - FrameLength);
            FOR i := 0 TO RemainBytes - 1 DO Rx[i] := Rx[TO_INT(FrameLength) + i]; END_FOR;
            RxCount := RxCount - FrameLength;
            FrameLength := 0;
            IF RxCount >= 7 THEN
                FrameLength := UDINT#6 + TO_UDINT(Rx[4])*256 + TO_UDINT(Rx[5]);
                IF (FrameLength < 9) OR (FrameLength > 260) THEN OperationFailed := TRUE; FailQuality := 'BAD_PROTOCOL';
                ELSIF RxCount >= FrameLength THEN State := 40;
                ELSE State := 30;
                END_IF;
            ELSE State := 30;
            END_IF;
        ELSE
            RxCount := 0; FrameLength := 0; State := 30;
        END_IF;
    ELSIF (RxCount = FrameLength) AND (FrameLength = UDINT#9)
        AND (Rx[0] = Tx[0]) AND (Rx[1] = Tx[1])
        AND (Rx[2] = BYTE#0) AND (Rx[3] = BYTE#0)
        AND (Rx[6] = Tx[6]) AND (Rx[7] = (FunctionCode OR BYTE#16#80))
        AND BlockHasHoles THEN
        (* Slave rejected a hole-bridged read with Modbus Exception: fall back to contiguous reads. *)
        HoleMergeDisabled := TRUE;
        FOR k := 2 TO BlockCount DO
            CandIndex := BlockIndices[k];
            Buffer.Cursors[CandIndex].NextDueMonoMs := SavedNextDue[k];
            Samples[CandIndex].NextPollMs := SavedNextDue[k];
        END_FOR;
        Point := Points[BlockIndices[1]];
        Width := UINT#1;
        IF (Point.dataType = 'float32') OR (Point.dataType = 'int32') OR (Point.dataType = 'uint32') THEN Width := UINT#2; END_IF;
        BlockCount := 1;
        BlockStartAddr := Point.address;
        BlockEndAddr := Point.address + Width;
        BlockWidth := Width;
        BlockHasHoles := FALSE;
        Retry := USINT#0;
        StaleDrains := USINT#0;
        State := 18;
    ELSIF (RxCount <> FrameLength) OR (Rx[0] <> Tx[0]) OR (Rx[1] <> Tx[1]) OR (Rx[2] <> 0) OR (Rx[3] <> 0) OR (Rx[6] <> Tx[6]) OR (Rx[7] <> FunctionCode) THEN
        OperationFailed := TRUE; FailQuality := 'BAD_PROTOCOL';
    ELSE
        IF Point.dataType = 'bool' THEN ByteCount := UINT#1; ELSE ByteCount := BlockWidth * UINT#2; END_IF;
        IF (TO_UINT(Rx[8]) <> ByteCount) OR (FrameLength <> TO_UDINT(UINT#9+ByteCount)) THEN OperationFailed := TRUE; FailQuality := 'BAD_PROTOCOL';
        ELSE
            BackoffLevel := USINT#0;
            IF NowMs >= RequestSentMs THEN LastRttMs := NowMs - RequestSentMs; ELSE LastRttMs := ULINT#0; END_IF;
            IF InterFrameGapMs > UDINT#0 THEN
                NextTxAllowedMs := NowMs + TO_ULINT(InterFrameGapMs);
            ELSIF LastRttMs >= ULINT#150 THEN
                NextTxAllowedMs := NowMs + ULINT#150;
            ELSE
                NextTxAllowedMs := ULINT#0;
            END_IF;
            AnyGoodInBlock := FALSE;
            AnyErrorInBlock := FALSE;
            BlockLastErr := '';
            SourceMarkUs := GET_MICROSECONDS(TRUE);
            FOR k := 1 TO BlockCount DO
                CandIndex := BlockIndices[k];
                Point := Points[CandIndex];
                PointDecodeFailed := FALSE;
                Width := UINT#1;
                IF (Point.dataType = 'float32') OR (Point.dataType = 'int32') OR (Point.dataType = 'uint32') THEN Width := UINT#2; END_IF;
                IF Point.dataType = 'bool' THEN
                    IF (Rx[9] AND BYTE#1) <> 0 THEN Value := 1; ELSE Value := 0; END_IF;
                ELSE
                    RawOff := 9 + TO_INT(Point.address - BlockStartAddr) * 2;
                    Decode[0] := Rx[RawOff]; Decode[1] := Rx[RawOff + 1];
                    IF Width = UINT#2 THEN Decode[2] := Rx[RawOff + 2]; Decode[3] := Rx[RawOff + 3];
                    ELSE Decode[2] := BYTE#0; Decode[3] := BYTE#0; END_IF;
                    IF (Point.byteOrder = 'BA') OR (Point.byteOrder = 'BADC') OR (Point.byteOrder = 'DCBA') THEN
                        Decode[0] := Rx[RawOff + 1]; Decode[1] := Rx[RawOff];
                        IF Width = UINT#2 THEN Decode[2] := Rx[RawOff + 3]; Decode[3] := Rx[RawOff + 2]; END_IF;
                    END_IF;
                    IF (Point.byteOrder = 'CDAB') OR (Point.byteOrder = 'DCBA') THEN
                        IF Point.byteOrder = 'CDAB' THEN
                            Decode[0] := Rx[RawOff + 2]; Decode[1] := Rx[RawOff + 3]; Decode[2] := Rx[RawOff]; Decode[3] := Rx[RawOff + 1];
                        ELSE
                            Decode[0] := Rx[RawOff + 3]; Decode[1] := Rx[RawOff + 2]; Decode[2] := Rx[RawOff + 1]; Decode[3] := Rx[RawOff];
                        END_IF;
                    END_IF;
                    UIntValue := TO_UDINT(Decode[0])*256 + TO_UDINT(Decode[1]);
                    IF Width = UINT#2 THEN UIntValue := UIntValue*65536 + TO_UDINT(Decode[2])*256 + TO_UDINT(Decode[3]); END_IF;
                    IF Point.dataType = 'float32' THEN
                        IF (TO_DWORD(UIntValue) AND DWORD#16#7F800000) = DWORD#16#7F800000 THEN
                            PointDecodeFailed := TRUE;
                        ELSE
                            ToFloat(REQ := FALSE, BUF_FORMAT := TRUE, BUF_OFFS := 0, BUF_CNT := 4, BUFFER := Decode, DST := FloatValue);
                            ToFloat(REQ := TRUE, BUF_FORMAT := TRUE, BUF_OFFS := 0, BUF_CNT := 4, BUFFER := Decode, DST := FloatValue);
                            Value := TO_LREAL(FloatValue);
                        END_IF;
                    ELSE
                        IntValue := TO_LINT(UIntValue);
                        IF (Point.dataType = 'int16') AND (UIntValue >= 32768) THEN IntValue := IntValue - 65536; END_IF;
                        IF (Point.dataType = 'int32') AND (UIntValue >= UDINT#2147483648) THEN IntValue := IntValue - LINT#4294967296; END_IF;
                        Value := TO_LREAL(IntValue);
                    END_IF;
                END_IF;
                IF PointDecodeFailed THEN
                    SourceResult(Index:=CandIndex, Value:=LREAL#0.0, Quality:='BAD_DECODE', NowMs:=NowMs, UnixMs:=UnixMs, NominalDueMs:=BlockNominalDue[k], ConfigSlot:=RequestSlot, ConfigGeneration:=RequestConfigGeneration, SamplingGeneration:=RequestSamplingGeneration, Samples:=Samples, Buffer:=Buffer);
                    Accepted:=SourceResult.Accepted;
                    AnyErrorInBlock := TRUE; BlockLastErr := 'BAD_DECODE';
                ELSE
                    SourceResult(Index:=CandIndex, Value:=Value*Point.scale+Point.offset, Quality:='GOOD', NowMs:=NowMs, UnixMs:=UnixMs, NominalDueMs:=BlockNominalDue[k], ConfigSlot:=RequestSlot, ConfigGeneration:=RequestConfigGeneration, SamplingGeneration:=RequestSamplingGeneration, Samples:=Samples, Buffer:=Buffer);
                    Accepted:=SourceResult.Accepted;
                    IF Samples[CandIndex].Quality='GOOD' THEN AnyGoodInBlock := TRUE;
                    ELSE AnyErrorInBlock := TRUE; BlockLastErr := Samples[CandIndex].Quality; END_IF;
                END_IF;
                IF Completed<UDINT#4294967295 THEN Completed:=Completed+1; END_IF;
            END_FOR;
            Buffer.SourceWorkUs:=Buffer.SourceWorkUs+GET_MICROSECONDS(TRUE)-SourceMarkUs;
            IF AnyGoodInBlock THEN LastGoodTimestamp:=UnixMs; END_IF;
            IF AnyErrorInBlock THEN StateText:='DEGRADED'; LastError:=BlockLastErr;
            ELSE StateText:='ONLINE'; LastError:=''; END_IF;
            State:=15;
        END_IF;
    END_IF;
90:
    IF NOT Socket.ACTIVE AND NOT Socket.BUSY THEN
        IF Enable AND Device.enabled AND NOT Reset AND (NowMs >= RetryAt) THEN State := 0;
        ELSIF Enable AND Device.enabled THEN StateText := 'OFFLINE';
        ELSE StateText := 'DISABLED'; END_IF;
    END_IF;
END_CASE;
IF OperationFailed THEN
    TimeoutRetryCap := Device.retryCount;
    IF TimeoutRetryCap > MaxTimeoutRetries THEN TimeoutRetryCap := MaxTimeoutRetries; END_IF;
    CanRetry := ((FailQuality = 'BAD_PROTOCOL') AND (Retry < Device.retryCount))
        OR ((FailQuality = 'BAD_TIMEOUT') AND TimeoutInReceive AND Socket.ACTIVE AND (Retry < TimeoutRetryCap));
    IF CanRetry THEN
        Retry := Retry + USINT#1;
        IF (FailQuality = 'BAD_TIMEOUT') OR (LastRttMs >= ULINT#150) THEN
            IF InterFrameGapMs >= UDINT#200 THEN NextTxAllowedMs := NowMs + TO_ULINT(InterFrameGapMs);
            ELSE NextTxAllowedMs := NowMs + ULINT#200; END_IF;
            State := 16;
        ELSIF InterFrameGapMs > UDINT#0 THEN
            NextTxAllowedMs := NowMs + TO_ULINT(InterFrameGapMs);
            State := 16;
        ELSE
            State := 18;
        END_IF;
    ELSE
        SourceMarkUs:=GET_MICROSECONDS(TRUE);
        FOR k := 1 TO BlockCount DO
            CandIndex := BlockIndices[k];
            SourceResult(Index:=CandIndex, Value:=LREAL#0.0, Quality:=FailQuality, NowMs:=NowMs, UnixMs:=UnixMs, NominalDueMs:=BlockNominalDue[k], ConfigSlot:=RequestSlot, ConfigGeneration:=RequestConfigGeneration, SamplingGeneration:=RequestSamplingGeneration, Samples:=Samples, Buffer:=Buffer);
            Accepted:=SourceResult.Accepted;
        END_FOR;
        Buffer.SourceWorkUs:=Buffer.SourceWorkUs+GET_MICROSECONDS(TRUE)-SourceMarkUs;
        LastError := FailQuality; StateText := 'DEGRADED';
        IF (FailQuality = 'BAD_TIMEOUT') OR (FailQuality = 'BAD_CONNECTION') THEN
            IF BackoffLevel < USINT#5 THEN BackoffLevel := BackoffLevel + USINT#1; END_IF;
            BackoffMs := ULINT#1000;
            FOR i := 1 TO TO_INT(BackoffLevel) DO
                IF BackoffMs < ULINT#15000 THEN BackoffMs := BackoffMs * ULINT#2; ELSE BackoffMs := ULINT#30000; END_IF;
            END_FOR;
            StateText := 'OFFLINE';
            RetryAt := NowMs + BackoffMs + TO_ULINT(Device.unitId MOD USINT#8) * ULINT#125;
            State := 90;
        ELSE State := 15; END_IF;
    END_IF;
END_IF;
END_FUNCTION_BLOCK

(* ---- NG_Mqtt.st ---- *)
FUNCTION_BLOCK NG_Mqtt
VAR_INPUT
    Enable : BOOL;
    BootId : NG_Id;
    Reconnect : BOOL;
    NowMs : ULINT;
    Bootstrap : NG_Bootstrap;
    TxRequest : BOOL;
    TxTopic : STRING[200];
    TxLength : UDINT;
    TxRetain : BOOL;
    RxAccept : BOOL;
    PlatformTime : BOOL;
    TxKind : INT;
    TxClockRevision : ULINT;
    TxBootId : NG_Id;
    TxConnectionRevision : ULINT;
    ClockRevision : ULINT;
    ConnectionRevision : ULINT;
    SnapshotMonoMs : ULINT;
    ControlAllowed : BOOL;
    SendAllowed : BOOL;
    TimeRequestId : NG_Id;
END_VAR
VAR_IN_OUT
    TxBuffer : NG_Bytes;
    RxBuffer : NG_Bytes;
END_VAR
VAR_OUTPUT
    Connected : BOOL;
    TxBusy : BOOL;
    TxDone : BOOL;
    RxReady : BOOL;
    RxTopic : STRING[500];
    RxLength : UDINT;
    RxRetained : BOOL;
    ErrorText : NG_Text;
    SessionCount : UDINT;
    WillCapacity : UDINT;
    WillEnabled : BOOL;
    DebugState : INT;
    TxInvoked : BOOL;
    TxSubmitted : BOOL;
    TxRejected : BOOL;
    SubmittedKind : INT;
    TxSubmitMonoMs : ULINT;
    RxReceivedMonoMs : ULINT;
END_VAR
VAR
    Client : IIoT_MqttClient_6;
    Options : MQTT_UDT_CONNECT_OPTIONS;
    ConnectStatus : MQTT_UDT_METHOD_STATUS;
    ConsumeStatus : MQTT_UDT_METHOD_STATUS;
    SubscribeStatus : MQTT_UDT_METHOD_STATUS;
    PublishStatus : MQTT_UDT_METHOD_STATUS;
    ReceiveStatus : MQTT_UDT_METHOD_STATUS;
    CheckStatus : MQTT_UDT_METHOD_STATUS;
    Info : MQTT_UDT_MESSAGE_INFO;
    State : INT;
    SubscribeIndex : INT;
    Filter : STRING[200];
    Prefix : STRING[150];
    server : STRING[200];
    id : STRING[128];
    user : STRING;
    password : STRING;
    ReadyClient : BOOL;
    NewMessage : BOOL;
    ConnectedResult : BOOL;
    ConsumeReq : BOOL;
    CheckReq : BOOL;
    PublishReq : BOOL;
    LastCheck : ULINT;
    RetryAt : ULINT;
    Deadline : ULINT;
    PrevTx : BOOL;
    WillSession : NG_Id;
    WillPayload : STRING[512];
    PublishPulse : BOOL;
    PublishLength : UDINT;
    TimePayload : STRING[512];
    TimeCopy : STRING_TO_BUF;
    TimePermit : NG_TimePermit;
END_VAR
TxDone := FALSE;
TxInvoked:=FALSE; TxSubmitted:=FALSE; TxRejected:=FALSE;
IF RxAccept THEN RxReady := FALSE; END_IF;
IF Reconnect OR NOT Enable THEN State := 900; END_IF;
IF State = 0 THEN
    server := Bootstrap.BrokerUri; id := Bootstrap.ClientId;
    user := Bootstrap.UserName; password := Bootstrap.Password;
    Prefix := CONCAT('iot/v1/gateway/',Bootstrap.GatewayId,'/');
    Options.diConnectTimeout := 5; Options.diKeepAliveInterval := 20;
    Options.xCleanSession := TRUE; Options.diMqttVersion := 4;
    Options.diMaxInflight := 4; Options.xAutomaticReconnect := FALSE;
    WillSession:=CONCAT(BootId,'-',TO_STRING(SessionCount+1,'{0:d}'));
    WillCapacity:=80; (* Vendor field is IecString80; SIZEOF also includes terminator/header. *)
    WillPayload:=CONCAT('{"schemaVersion":1,"gatewayId":',NG_Quote(Bootstrap.GatewayId),',"timestamp":null,"sessionId":',NG_Quote(WillSession),',"online":false,"reason":"connection_lost"}');
    WillEnabled:=(TO_UDINT(LEN(WillPayload))<=WillCapacity) AND (LEN(Prefix)+6<=80);
    Options.xUseWillOptions:=WillEnabled;
    IF WillEnabled THEN
        Options.udtWill.strTopic:=CONCAT(Prefix,'status'); Options.udtWill.strPayload:=WillPayload;
    ELSE Options.udtWill.strTopic:=''; Options.udtWill.strPayload:=''; END_IF;
    Options.udtWill.diQos:=1; Options.udtWill.xRetained:=TRUE;
    ErrorText := ''; Connected := FALSE; Deadline := NowMs + 15000;
    State := 5;
END_IF;
Client(EN := Enable AND (State < 900), strServerUri := server, strClientId := id, strPersistDir := '', diMaxBufferedMessages := DINT#0, ENO => ReadyClient);
Client.Connect(State = 10, user, password, Options, ConnectStatus);
Client.StartConsuming(State = 20, ConsumeStatus);
Client.Subscribe(State = 30, Filter, DINT#1, SubscribeStatus);
(* This is the library request entry, one scan after Main's TxRequest.
   Encode m1 here so local publisher waiting is never excluded from RTT. *)
PublishPulse:=PublishReq;
IF PublishPulse AND PlatformTime THEN
    IF TxKind=8 THEN
        TxSubmitMonoMs:=NowMs;
        TimePayload:=CONCAT('{"schemaVersion":1,"gatewayId":',NG_Quote(Bootstrap.GatewayId),',"requestId":',NG_Quote(TimeRequestId),',"bootId":',NG_Quote(BootId),',"sessionId":',NG_Quote(WillSession),',"clientMonoMs":',TO_STRING(TxSubmitMonoMs,'{0:d}'),'}');
        TimeCopy(REQ:=FALSE,BUF_FORMAT:=FALSE,BUF_OFFS:=0,BUF_CNT:=LEN(TimePayload),SRC:=TimePayload,BUFFER:=TxBuffer);
        TimeCopy(REQ:=TRUE,BUF_FORMAT:=FALSE,BUF_OFFS:=0,BUF_CNT:=LEN(TimePayload),SRC:=TimePayload,BUFFER:=TxBuffer);
        PublishPulse:=TimeCopy.DONE AND NG_ValidId(TimeRequestId) AND (NowMs<=ULINT#9007199254740991);
    ELSE
        TimePermit(Purpose:=USINT#3,TokenBootId:=TxBootId,CurrentBootId:=BootId,NowMs:=NowMs,TokenMonoMs:=SnapshotMonoMs,
            TokenClockRevision:=TxClockRevision,TokenConnectionRevision:=TxConnectionRevision,
            CurrentClockRevision:=ClockRevision,CurrentConnectionRevision:=ConnectionRevision,
            EnqueueAllowed:=FALSE,ControlAllowed:=ControlAllowed,SendAllowed:=SendAllowed,AckApplyAllowed:=Connected);
        PublishPulse:=TimePermit.Allowed;
        IF (TxKind=5) OR (TxKind=6) THEN PublishPulse:=PublishPulse AND SendAllowed; END_IF;
    END_IF;
    IF NOT PublishPulse THEN TxRejected:=TRUE; TxBusy:=FALSE; END_IF;
END_IF;
IF PublishPulse AND (TxKind=5) AND NOT SendAllowed THEN
    PublishPulse:=FALSE; TxRejected:=TRUE; TxBusy:=FALSE;
END_IF;
IF PublishPulse THEN TxInvoked:=TRUE; TxSubmitMonoMs:=NowMs; SubmittedKind:=TxKind; END_IF;
PublishLength:=TxLength;
IF PlatformTime AND (TxKind=8) THEN PublishLength:=TO_UDINT(LEN(TimePayload)); END_IF;
Client.Publish(PublishPulse,TxTopic,TxBuffer,PublishLength,DINT#1,TxRetain,PublishStatus);
IF PublishPulse THEN
    (* Busy proves the asynchronous method accepted the request. Done is also
       sufficient; no PUBACK is required to create the Busy submission fact. *)
    TxSubmitted:=NOT PublishStatus.xError AND (PublishStatus.xBusy OR PublishStatus.xDone);
    IF PublishStatus.xError THEN TxRejected:=TRUE; TxBusy:=FALSE; END_IF;
END_IF;
NewMessage := Client.TryConsumeMessage(ConsumeReq, RxTopic, RxBuffer, Info, ReceiveStatus);
ConnectedResult := Client.IsConnected(CheckReq, CheckStatus);
PublishReq := FALSE;
CASE State OF
5:
    IF Client.xError THEN ErrorText := 'MQTT_CLIENT_ERROR'; State := 900;
    ELSIF ReadyClient THEN State := 10;
    END_IF;
10: State := 11;
11:
    IF ConnectStatus.xError THEN ErrorText := 'MQTT_CONNECT_ERROR'; State := 900;
    ELSIF ConnectStatus.xDone THEN State := 20; END_IF;
20: State := 21;
21:
    IF ConsumeStatus.xError THEN ErrorText := 'MQTT_CONSUME_ERROR'; State := 900;
    ELSIF ConsumeStatus.xDone THEN SubscribeIndex := 1; State := 25; END_IF;
25:
    CASE SubscribeIndex OF
        1: Filter := CONCAT(Prefix,'config/set');
        2: Filter := CONCAT(Prefix,'config/patch');
        3: Filter := CONCAT(Prefix,'data/ack');
        4: Filter := CONCAT(Prefix,'time/response');
    END_CASE;
    State := 30;
30: State := 31;
31:
    IF SubscribeStatus.xError THEN ErrorText := 'MQTT_SUBSCRIBE_ERROR'; State := 900;
    ELSIF SubscribeStatus.xDone THEN
        IF (SubscribeIndex < 3) OR (PlatformTime AND (SubscribeIndex<4)) THEN SubscribeIndex := SubscribeIndex+1; State := 25;
        ELSE Connected := TRUE; ErrorText := ''; SessionCount := SessionCount+1; State := 100; END_IF;
    END_IF;
100:
    IF TxRequest AND NOT PrevTx AND NOT TxBusy THEN TxBusy := TRUE; PublishReq := TRUE; END_IF;
    IF TxBusy THEN
        IF PublishStatus.xDone THEN TxBusy := FALSE; TxDone := TRUE;
        ELSIF PublishStatus.xError THEN ErrorText := 'MQTT_PUBLISH_ERROR'; State := 900; END_IF;
    END_IF;
    IF NOT RxReady THEN
        IF ReceiveStatus.xDone THEN
            IF NewMessage THEN
                RxLength := Info.udiLength; RxRetained := Info.xRetained; RxReady := TRUE;
                (* Earliest ST-visible receive boundary. Queue/scan delay remains
                   inside complete request-to-dequeue RTT and asymmetry bound. *)
                RxReceivedMonoMs:=NowMs;
            END_IF;
            ConsumeReq := FALSE;
        ELSIF NOT ReceiveStatus.xBusy THEN ConsumeReq := NOT ConsumeReq; END_IF;
    ELSE ConsumeReq := FALSE;
    END_IF;
    IF ReceiveStatus.xError THEN
        (* Hub clears retained config/set with a zero-byte publication before a patch.
           IIoT 5.3 reports this as diagnostic 10 / Null message received. Keep
           consuming so the following patch is preserved; IsConnected still
           detects a real connection loss. All other receive errors reconnect. *)
        IF NOT ((ReceiveStatus.udtDiag.wDiagCode=WORD#10) AND
                (ReceiveStatus.udtDiag.strDiagMsg='Null message received')) THEN
            ErrorText := CONCAT('MQTT_RECEIVE_ERROR: ',ReceiveStatus.udtDiag.strDiagMsg); State := 900;
        END_IF;
    END_IF;
    IF CheckStatus.xDone THEN
        CheckReq := FALSE; LastCheck := NowMs;
        IF NOT ConnectedResult THEN ErrorText := 'MQTT_DISCONNECTED'; State := 900; END_IF;
    ELSIF (NowMs > LastCheck + 2000) AND NOT CheckStatus.xBusy THEN CheckReq := TRUE; END_IF;
900:
    Connected := FALSE; TxBusy := FALSE; ConsumeReq := FALSE; CheckReq := FALSE; PublishReq := FALSE;
    RetryAt := NowMs + 3000; State := 910;
910:
    IF NOT ReadyClient AND NOT Client.xBusy AND Enable AND NOT Reconnect AND (NowMs >= RetryAt) THEN State := 0; END_IF;
END_CASE;
IF (State > 0) AND (State < 100) AND (NowMs >= Deadline) THEN ErrorText := 'MQTT_TIMEOUT'; State := 900; END_IF;
PrevTx := TxRequest;
DebugState:=State;
END_FUNCTION_BLOCK

(* ---- NG_PlatformTime.st ---- *)
FUNCTION_BLOCK NG_PlatformTime
VAR_INPUT
    Reset : BOOL;
    PlatformMode : BOOL;
    Connected : BOOL;
    SessionId : NG_Id;
    NowMs : ULINT;
    SystemUtcMs : ULINT;
    TimeBasisRef : NG_Id;
    DriftBoundPpm : LREAL;
    DriftEvidence : NG_Text;
    HistoryBasisRef : NG_Id;
    HistoryUtcLowerMs : ULINT;
    RequestSubmitted : BOOL;
    RequestSubmittedMonoMs : ULINT;
    ResponseReady : BOOL;
    ResponseClientMonoMs : ULINT;
    ResponseReceivedMonoMs : ULINT;
    ServerReceivedMs : ULINT;
    ServerSentMs : ULINT;
    HeartbeatSubmitted : BOOL;
    ConfigGetSubmitted : BOOL;
END_VAR
VAR_OUTPUT
    State : USINT;
    TimeValid : BOOL;
    UtcMs : ULINT;
    UncertaintyMs : ULINT;
    SyncAgeMs : ULINT;
    ClockRevision : ULINT;
    ConnectionRevision : ULINT;
    CaptureAllowed : BOOL;
    EnqueueAllowed : BOOL;
    ControlAllowed : BOOL;
    SendAllowed : BOOL;
    AckApplyAllowed : BOOL;
    RequestWanted : BOOL;
    RequestId : NG_Id;
    RequestClientMonoMs : ULINT;
    PendingRequest : BOOL;
    Attempts : UINT;
    HeartbeatReady : BOOL;
    ConfigGetReady : BOOL;
    ErrorText : NG_Text;
END_VAR
VAR
    Started : BOOL;
    SeenConnected : BOOL;
    SeenSession : NG_Id;
    SeenPlatformMode : BOOL;
    SeenBasis : NG_Id;
    SeenDrift : LREAL;
    SeenDriftEvidence : NG_Text;
    SessionChecked : BOOL;
    HeartbeatAccepted : BOOL;
    GetAccepted : BOOL;
    LastMono : ULINT;
    Anchor : LREAL;
    HasAnchor : BOOL;
    Residual : LREAL;
    BaseError : LREAL;
    LastSync : ULINT;
    RoundStart : ULINT;
    RoundOpen : BOOL;
    NextSync : ULINT;
    Failures : UINT;
    RequestSequence : ULINT;
    Candidates : UINT;
    CandidateUtc : ARRAY[1..3] OF LREAL;
    CandidateMono : ARRAY[1..3] OF ULINT;
    CandidatePath : ARRAY[1..3] OF LREAL;
    CandidateError : ARRAY[1..3] OF LREAL;
    CandidateRtt : ARRAY[1..3] OF ULINT;
    ConfirmDeviation : BOOL;
    Elapsed : LREAL;
    Correction : LREAL;
    ErrorBound : LREAL;
    Rtt : LREAL;
    Processing : LREAL;
    PathMs : LREAL;
    Target : LREAL;
    CandidateLow : LREAL;
    CandidateHigh : LREAL;
    ChosenError : LREAL;
    PreviousError : LREAL;
    RecoveryTolerance : LREAL;
    OutputFloor : LREAL;
    LastOutputUtc : ULINT;
    BestPath : LREAL;
    DelayMs : ULINT;
    FinishRound : BOOL;
    Adopt : BOOL;
    Invalidate : BOOL;
    WasValid : BOOL;
    Chosen : UINT;
    i : UINT;
END_VAR
(* Pure clock kernel: no RTC writes, file, socket, device or vendor timing calls.
   ResponseReady must come from NG_TimeResponse after exact echo/retained checks.
   RequestSubmitted/control inputs mean synchronous SDK acceptance, never PUBACK.
   State: 0 UNSYNCED, 1 SYNCING, 2 SYNCED, 3 HOLDOVER, 4 EXPIRED,
          5 SUSPECT, 6 MAINTENANCE. Reset means a NEW boot only. *)
IF Reset OR NOT Started THEN
    Started:=TRUE; State:=0; HasAnchor:=FALSE; TimeValid:=FALSE; Anchor:=0;
    Residual:=0; ClockRevision:=0; ConnectionRevision:=0; LastMono:=NowMs;
    SeenConnected:=FALSE; SeenSession:=''; SessionChecked:=FALSE;
    SeenPlatformMode:=PlatformMode; SeenBasis:=TimeBasisRef;
    SeenDrift:=DriftBoundPpm; SeenDriftEvidence:=DriftEvidence;
    HeartbeatAccepted:=FALSE; GetAccepted:=FALSE; PendingRequest:=FALSE;
    RequestWanted:=FALSE; RoundOpen:=FALSE; NextSync:=0; RequestSequence:=0;
    Attempts:=0; Candidates:=0; Failures:=0; ConfirmDeviation:=FALSE; ErrorText:='';
    LastOutputUtc:=0;
END_IF;
WasValid:=TimeValid; Invalidate:=FALSE; Adopt:=FALSE; FinishRound:=FALSE;
IF (PlatformMode<>SeenPlatformMode) OR (TimeBasisRef<>SeenBasis)
    OR (DriftBoundPpm<>SeenDrift) OR (DriftEvidence<>SeenDriftEvidence) THEN
    State:=6; Invalidate:=TRUE; ErrorText:='TIME_SOURCE_CHANGE_REQUIRES_MAINTENANCE';
END_IF;
IF NowMs<LastMono THEN
    State:=6; HasAnchor:=FALSE; Invalidate:=TRUE; ErrorText:='CLOCK_CONTINUITY_REQUIRES_MAINTENANCE';
END_IF;
Elapsed:=0; IF NowMs>=LastMono THEN Elapsed:=TO_LREAL(NowMs-LastMono); END_IF;
IF HasAnchor THEN
    Correction:=MAX(-Elapsed*LREAL#0.005,MIN(Elapsed*LREAL#0.005,Residual));
    Anchor:=Anchor+Elapsed+Correction; Residual:=Residual-Correction;
END_IF;
LastMono:=NowMs;
IF (Connected<>SeenConnected) OR (Connected AND (SessionId<>SeenSession)) THEN
    IF ConnectionRevision>=ULINT#9007199254740991 THEN State:=6; ErrorText:='CONNECTION_REVISION_EXHAUSTED';
    ELSE ConnectionRevision:=ConnectionRevision+1; END_IF;
    SeenConnected:=Connected; SeenSession:=SessionId; SessionChecked:=FALSE;
    HeartbeatAccepted:=FALSE; GetAccepted:=FALSE; PendingRequest:=FALSE;
    RequestWanted:=FALSE; RoundOpen:=FALSE; Candidates:=0; Attempts:=0; NextSync:=NowMs;
END_IF;
IF PlatformMode THEN
    IF NOT NG_ValidId(TimeBasisRef) OR (DriftEvidence='') OR NOT ((DriftBoundPpm>=0) AND (DriftBoundPpm<=1000)) THEN
        State:=6; Invalidate:=TRUE; ErrorText:='MISSING_TIME_BASIS_OR_DRIFT_EVIDENCE';
    END_IF;
    IF (HistoryUtcLowerMs>0) AND (HistoryBasisRef<>TimeBasisRef) THEN
        State:=6; Invalidate:=TRUE; ErrorText:='HISTORY_BASIS_REQUIRES_MAINTENANCE';
    END_IF;
    IF PendingRequest AND (NowMs>=RequestClientMonoMs+2000) THEN PendingRequest:=FALSE; END_IF;
    IF ResponseReady AND PendingRequest AND (State<>6) THEN
        (* Reader is required to compare the exact six request fields first. *)
        PendingRequest:=FALSE;
        IF (ResponseClientMonoMs=RequestClientMonoMs) AND (ResponseReceivedMonoMs>=RequestClientMonoMs)
            AND (ResponseReceivedMonoMs<=NowMs) AND (NowMs<RequestClientMonoMs+2000)
            AND (ServerSentMs>=ServerReceivedMs) AND (ServerSentMs<=ULINT#9007199254740991) THEN
            Rtt:=TO_LREAL(ResponseReceivedMonoMs-RequestClientMonoMs);
            Processing:=TO_LREAL(ServerSentMs-ServerReceivedMs); PathMs:=Rtt-Processing;
            Target:=TO_LREAL(ServerSentMs)+MAX(LREAL#0.0,PathMs)/2;
            ErrorBound:=MAX(LREAL#0.0,PathMs)/2+MAX(LREAL#0.0,-PathMs)+22;
            IF (Rtt<2000) AND (Processing<=500) AND (PathMs>=-50)
                AND (Target-ErrorBound>=0) AND (Target+ErrorBound<=LREAL#9007199254740991.0) THEN
                IF Candidates<3 THEN
                    Candidates:=Candidates+1; CandidateUtc[Candidates]:=Target;
                    CandidateMono[Candidates]:=ResponseReceivedMonoMs; CandidatePath[Candidates]:=MAX(LREAL#0.0,PathMs);
                    CandidateError[Candidates]:=ErrorBound; CandidateRtt[Candidates]:=TO_ULINT(Rtt);
                    IF Candidates=3 THEN FinishRound:=TRUE; END_IF;
                END_IF;
            ELSE ErrorText:='HIGH_DELAY_OR_UNSAFE_TIME'; END_IF;
        ELSE ErrorText:='STALE_TIME_RESPONSE'; END_IF;
    END_IF;
    IF RoundOpen AND ((NowMs>=RoundStart+30000) OR ((Attempts>=10) AND NOT PendingRequest)) THEN FinishRound:=TRUE; END_IF;
    IF FinishRound THEN
        Chosen:=0; CandidateLow:=LREAL#9007199254740991.0; CandidateHigh:=0; BestPath:=LREAL#9007199254740991.0;
        FOR i:=1 TO Candidates DO
            Target:=CandidateUtc[i]+TO_LREAL(NowMs-CandidateMono[i]);
            CandidateLow:=MIN(CandidateLow,Target); CandidateHigh:=MAX(CandidateHigh,Target);
            IF ((Candidates>=3) OR (CandidateRtt[i]<=500)) AND (CandidatePath[i]<BestPath) THEN
                Chosen:=i; BestPath:=CandidatePath[i];
            END_IF;
        END_FOR;
        IF (Chosen>0) AND (CandidateHigh-CandidateLow<=500) THEN
            Target:=CandidateUtc[Chosen]+TO_LREAL(NowMs-CandidateMono[Chosen]);
            ChosenError:=CandidateError[Chosen]+TO_LREAL(NowMs-CandidateMono[Chosen])*DriftBoundPpm/LREAL#1000000.0;
            (* A holdover estimate is not a timestamp already emitted. Include
               its accumulated drift error before declaring a discontinuity.
               Larger changes need a second consistent round, never a latch
               which prevents the next time request. Output remains monotonic. *)
            PreviousError:=0;
            IF HasAnchor THEN PreviousError:=BaseError+TO_LREAL(NowMs-LastSync)*DriftBoundPpm/LREAL#1000000.0+ABS(Residual); END_IF;
            RecoveryTolerance:=MAX(LREAL#5000.0,PreviousError+ChosenError);
            IF HasAnchor AND (ABS(Target-Anchor)>RecoveryTolerance) AND NOT ConfirmDeviation THEN
                State:=5; Invalidate:=TRUE; ErrorText:='TIME_CORRECTION_CONFIRMING';
                ConfirmDeviation:=TRUE; NextSync:=NowMs+10000;
            ELSE Adopt:=TRUE; END_IF;
            IF Adopt THEN
                OutputFloor:=MAX(TO_LREAL(LastOutputUtc),TO_LREAL(HistoryUtcLowerMs));
                IF NOT HasAnchor OR (State=4) OR (State=5) OR (State=0) OR (State=1) THEN
                    Anchor:=MAX(Target,OutputFloor); Residual:=Target-Anchor; HasAnchor:=TRUE;
                    IF ClockRevision>=ULINT#9007199254740991 THEN State:=6; Invalidate:=TRUE;
                    ELSE ClockRevision:=ClockRevision+1; END_IF;
                ELSE Residual:=Target-Anchor; END_IF;
                IF State<>6 THEN
                    BaseError:=ChosenError; LastSync:=NowMs; State:=2; SessionChecked:=Connected;
                    ConfirmDeviation:=FALSE; Failures:=0; ErrorText:=''; Invalidate:=FALSE;
                    IF Candidates<3 THEN NextSync:=NowMs+10000;
                    ELSE NextSync:=NowMs+270000+(RequestSequence MOD 60001); END_IF;
                END_IF;
            END_IF;
        ELSE
            Failures:=MIN(Failures+1,UINT#5); DelayMs:=5000;
            CASE Failures OF 2: DelayMs:=10000; 3: DelayMs:=20000; 4: DelayMs:=40000; 5: DelayMs:=60000; END_CASE;
            NextSync:=NowMs+MIN(ULINT#60000,DelayMs+(RequestSequence MOD 1001)); ErrorText:='TIMEOUT_OR_INCONSISTENT';
        END_IF;
        RoundOpen:=FALSE; PendingRequest:=FALSE; Candidates:=0;
    END_IF;
    IF (State<>6) AND Connected AND (NowMs>=NextSync) AND NOT PendingRequest THEN
        IF NOT RoundOpen THEN
            RoundOpen:=TRUE; RoundStart:=NowMs; Attempts:=0; Candidates:=0;
            IF NOT HasAnchor THEN State:=1; END_IF;
        END_IF;
        RequestWanted:=(Attempts<10) AND (NowMs<RoundStart+30000);
    ELSE RequestWanted:=FALSE; END_IF;
    IF RequestWanted THEN RequestId:=CONCAT('t-',TO_STRING(ConnectionRevision,'{0:d}'),'-',TO_STRING(RequestSequence+1,'{0:d}')); END_IF;
    IF RequestSubmitted AND RequestWanted THEN
        IF RequestSequence>=ULINT#9007199254740990 THEN State:=6; Invalidate:=TRUE; ErrorText:='REQUEST_SEQUENCE_EXHAUSTED';
        ELSE
            RequestSequence:=RequestSequence+1; RequestClientMonoMs:=NowMs;
            IF (RequestSubmittedMonoMs>0) AND (RequestSubmittedMonoMs<=NowMs) THEN RequestClientMonoMs:=RequestSubmittedMonoMs; END_IF;
            Attempts:=Attempts+1; PendingRequest:=TRUE; RequestWanted:=FALSE;
        END_IF;
    END_IF;
END_IF;
UtcMs:=0; UncertaintyMs:=0; SyncAgeMs:=0; TimeValid:=FALSE;
IF HasAnchor THEN
    SyncAgeMs:=NowMs-LastSync;
    ErrorBound:=BaseError+TO_LREAL(SyncAgeMs)*DriftBoundPpm/LREAL#1000000.0+ABS(Residual);
    (* Round up positive error; TO_ULINT rounds rather than truncates on target. *)
    IF (ErrorBound>=0) AND (ErrorBound<LREAL#9007199254740990.0) THEN
        UncertaintyMs:=TO_ULINT(TRUNC_LINT(ErrorBound));
        IF TO_LREAL(UncertaintyMs)<ErrorBound THEN UncertaintyMs:=UncertaintyMs+1; END_IF;
    END_IF;
    TimeValid:=PlatformMode AND ((State=2) OR (State=3)) AND (SyncAgeMs<3600000)
        AND (ErrorBound>=0) AND (UncertaintyMs<5000) AND (Anchor-ErrorBound>=0)
        AND (Anchor+ErrorBound<=LREAL#9007199254740991.0);
    IF TimeValid THEN
        UtcMs:=MAX(LastOutputUtc,TO_ULINT(TRUNC_LINT(Anchor))); LastOutputUtc:=UtcMs;
        IF SessionChecked THEN State:=2; ELSE State:=3; END_IF;
    ELSIF (State=2) OR (State=3) THEN
        State:=4; Invalidate:=TRUE;
        IF ABS(Residual)>=5000 THEN ErrorText:='TIME_CORRECTION_WAITING'; NextSync:=MIN(NextSync,NowMs+10000);
        ELSE ErrorText:='HOLDOVER_EXPIRED'; END_IF;
    END_IF;
END_IF;
IF Invalidate THEN
    IF WasValid THEN
        IF ClockRevision>=ULINT#9007199254740991 THEN State:=6;
        ELSE ClockRevision:=ClockRevision+1; END_IF;
    END_IF;
    SessionChecked:=FALSE; HeartbeatAccepted:=FALSE; GetAccepted:=FALSE;
END_IF;
CaptureAllowed:=TRUE; AckApplyAllowed:=Connected;
EnqueueAllowed:=TimeValid; ControlAllowed:=TimeValid AND Connected AND SessionChecked;
IF NOT PlatformMode AND (State<>6) THEN
    EnqueueAllowed:=(SystemUtcMs>0) AND (SystemUtcMs<=ULINT#9007199254740991);
    ControlAllowed:=EnqueueAllowed AND Connected; UtcMs:=SystemUtcMs;
END_IF;
IF ControlAllowed THEN
    IF HeartbeatSubmitted THEN HeartbeatAccepted:=TRUE; END_IF;
    IF ConfigGetSubmitted AND HeartbeatAccepted THEN GetAccepted:=TRUE; END_IF;
END_IF;
SendAllowed:=ControlAllowed AND HeartbeatAccepted AND GetAccepted;
HeartbeatReady:=HeartbeatAccepted; ConfigGetReady:=GetAccepted;
END_FUNCTION_BLOCK

(* ---- NG_PlatformTimeChecks.st ---- *)
FUNCTION_BLOCK NG_PlatformTimeChecks
VAR_OUTPUT
    Done : BOOL;
    Passed : UINT;
    FailedChecks : UINT;
    WirePassed : UINT;
    WireFailed : UINT;
END_VAR
VAR_IN_OUT
    Doc : NG_Document;
    Bytes : NG_Bytes;
END_VAR
VAR
    LogicalClock : NG_PlatformTime;
    Permit : NG_TimePermit;
    WireTests : NG_TimeResponseChecks;
    ClockDone : BOOL;
    Stage : UINT;
    Checks : ARRAY[1..40] OF BOOL;
    Tick : ULINT := 100000;
    ResetClock : BOOL;
    Connected : BOOL := TRUE;
    Session : NG_Id := 'session-one';
    Submit : BOOL;
    Reply : BOOL;
    Heartbeat : BOOL;
    GetConfig : BOOL;
    RequestMono : ULINT;
    ServerT3 : ULINT;
    SystemDate : ULINT := 1000;
    SavedClockRevision : ULINT;
    SavedConnectionRevision : ULINT;
    SavedOutput : ULINT;
    Drift : LREAL := 50;
    i : UINT;
END_VAR

(* Offline assertion program. No gateway, socket, store, physical IO or RTC writes.
   Cold compilation is not execution; Done/Checks need a later authorized test runtime. *)
WireTests(Doc:=Doc,Bytes:=Bytes);
WirePassed:=WireTests.Passed; WireFailed:=WireTests.FailedChecks;
Done:=ClockDone AND WireTests.Done;
IF ClockDone THEN RETURN; END_IF;
ResetClock:=FALSE; Submit:=FALSE; Reply:=FALSE; Heartbeat:=FALSE; GetConfig:=FALSE;
CASE Stage OF
    0: ResetClock:=TRUE;
    1,3,5: Submit:=TRUE; RequestMono:=Tick;
    2,4,6: Tick:=Tick+20; Reply:=TRUE; ServerT3:=ULINT#1792000000000+Tick-100000-9;
    7: GetConfig:=TRUE;
    8: Heartbeat:=TRUE;
    9: GetConfig:=TRUE;
    10: SystemDate:=ULINT#9000000000000; Tick:=Tick+20;
    11: Connected:=FALSE; Tick:=Tick+20;
    12: Connected:=TRUE; Session:='session-two'; Tick:=Tick+20;
    13: Tick:=Tick+3600000;
    14: Tick:=Tick-1;
    15: ResetClock:=TRUE; Tick:=100000; Drift:=1000; Session:='recover-one';
    16,18,20,24,26,28,33,35,37,40,42,44,47,49,51,54,56,58: Submit:=TRUE; RequestMono:=Tick;
    17,19,21: Tick:=Tick+20; Reply:=TRUE; ServerT3:=ULINT#1792000000000+Tick-100000-9;
    22: SavedOutput:=LogicalClock.UtcMs; Connected:=FALSE; Tick:=Tick+172800000;
    23: Connected:=TRUE; Session:='recover-two';
    25,27,29: Tick:=Tick+20; Reply:=TRUE; ServerT3:=ULINT#1792000000000+Tick-100000-9-2170;
    30,60: Heartbeat:=TRUE;
    31,61: GetConfig:=TRUE;
    32,39: Tick:=Tick+330000;
    34,36,38: Tick:=Tick+20; Reply:=TRUE; ServerT3:=ULINT#1792000000000+Tick-100000-9-4340;
    41,43,45,48,50,52,55,57,59: Tick:=Tick+20; Reply:=TRUE; ServerT3:=ULINT#1792000000000+Tick-100000-9-90000;
    46: Tick:=Tick+10000;
    53: Tick:=Tick+120000;
END_CASE;
IF (Stage=37) OR (Stage=44) THEN SavedOutput:=LogicalClock.UtcMs; END_IF;
LogicalClock(Reset:=ResetClock,PlatformMode:=TRUE,Connected:=Connected,SessionId:=Session,NowMs:=Tick,SystemUtcMs:=SystemDate,
    TimeBasisRef:='site-hub-1',DriftBoundPpm:=Drift,DriftEvidence:='TEST_FIXTURE_ONLY',HistoryBasisRef:='',HistoryUtcLowerMs:=0,
    RequestSubmitted:=Submit,ResponseReady:=Reply,ResponseClientMonoMs:=RequestMono,ResponseReceivedMonoMs:=Tick,
    ServerReceivedMs:=ServerT3-2,ServerSentMs:=ServerT3,HeartbeatSubmitted:=Heartbeat,ConfigGetSubmitted:=GetConfig);
CASE Stage OF
0:
    Checks[1]:=LogicalClock.CaptureAllowed AND LogicalClock.AckApplyAllowed AND NOT LogicalClock.EnqueueAllowed AND NOT LogicalClock.ControlAllowed;
    Checks[2]:=LogicalClock.RequestWanted AND NOT LogicalClock.TimeValid;
1: Checks[3]:=LogicalClock.PendingRequest AND (LogicalClock.RequestClientMonoMs=Tick) AND (LogicalClock.Attempts=1);
2: Checks[4]:=NOT LogicalClock.TimeValid AND LogicalClock.RequestWanted;
6:
    Checks[5]:=LogicalClock.TimeValid AND LogicalClock.ControlAllowed AND NOT LogicalClock.SendAllowed;
    Checks[6]:=(LogicalClock.UtcMs=ULINT#1792000000060) AND (LogicalClock.UncertaintyMs=32);
    SavedClockRevision:=LogicalClock.ClockRevision; SavedConnectionRevision:=LogicalClock.ConnectionRevision;
7: Checks[7]:=NOT LogicalClock.SendAllowed;
8: Checks[8]:=NOT LogicalClock.SendAllowed;
9: Checks[9]:=LogicalClock.SendAllowed;
10: Checks[10]:=LogicalClock.TimeValid AND (LogicalClock.UtcMs=ULINT#1792000000080);
11: Checks[11]:=LogicalClock.TimeValid AND LogicalClock.EnqueueAllowed AND NOT LogicalClock.ControlAllowed AND NOT LogicalClock.SendAllowed;
12:
    Checks[12]:=LogicalClock.TimeValid AND NOT LogicalClock.ControlAllowed AND NOT LogicalClock.SendAllowed;
    Checks[13]:=(LogicalClock.ClockRevision=SavedClockRevision) AND (LogicalClock.ConnectionRevision>SavedConnectionRevision);
    Permit(Purpose:=USINT#4,TokenBootId:='boot-one',CurrentBootId:='boot-one',NowMs:=Tick,TokenMonoMs:=Tick,
        TokenClockRevision:=SavedClockRevision,TokenConnectionRevision:=SavedConnectionRevision,
        CurrentClockRevision:=LogicalClock.ClockRevision,CurrentConnectionRevision:=LogicalClock.ConnectionRevision,
        EnqueueAllowed:=TRUE,ControlAllowed:=TRUE,SendAllowed:=TRUE,AckApplyAllowed:=TRUE);
    Checks[14]:=NOT Permit.Allowed;
13:
    Checks[15]:=NOT LogicalClock.TimeValid AND NOT LogicalClock.EnqueueAllowed AND LogicalClock.CaptureAllowed AND LogicalClock.AckApplyAllowed;
    Checks[16]:=LogicalClock.State=4;
14:
    Checks[17]:=(LogicalClock.State=6) AND NOT LogicalClock.TimeValid;
    Permit(Purpose:=USINT#5,TokenBootId:='',CurrentBootId:='boot-one',NowMs:=Tick,TokenMonoMs:=0,
        TokenClockRevision:=0,TokenConnectionRevision:=0,CurrentClockRevision:=99,CurrentConnectionRevision:=99,
        EnqueueAllowed:=FALSE,ControlAllowed:=FALSE,SendAllowed:=FALSE,AckApplyAllowed:=TRUE);
    Checks[18]:=Permit.Allowed;
    Permit(Purpose:=USINT#2,TokenBootId:='old-boot',CurrentBootId:='boot-one',NowMs:=Tick,TokenMonoMs:=Tick,
        TokenClockRevision:=0,TokenConnectionRevision:=0,CurrentClockRevision:=0,CurrentConnectionRevision:=0,
        EnqueueAllowed:=TRUE,ControlAllowed:=TRUE,SendAllowed:=TRUE,AckApplyAllowed:=TRUE);
    Checks[19]:=NOT Permit.Allowed;
    Permit(Purpose:=USINT#2,TokenBootId:='boot-one',CurrentBootId:='boot-one',NowMs:=Tick,TokenMonoMs:=Tick-2000,
        TokenClockRevision:=0,TokenConnectionRevision:=0,CurrentClockRevision:=0,CurrentConnectionRevision:=0,
        EnqueueAllowed:=TRUE,ControlAllowed:=TRUE,SendAllowed:=TRUE,AckApplyAllowed:=TRUE);
    Checks[20]:=NOT Permit.Allowed;
    Permit(Purpose:=USINT#2,TokenBootId:='boot-one',CurrentBootId:='boot-one',NowMs:=Tick,TokenMonoMs:=Tick,
        TokenClockRevision:=0,TokenConnectionRevision:=0,CurrentClockRevision:=0,CurrentConnectionRevision:=0,
        EnqueueAllowed:=TRUE,ControlAllowed:=TRUE,SendAllowed:=TRUE,AckApplyAllowed:=TRUE);
    Checks[21]:=Permit.Allowed;
    LogicalClock(Reset:=TRUE,PlatformMode:=FALSE,Connected:=TRUE,SessionId:='compat',NowMs:=Tick,SystemUtcMs:=SystemDate,
        TimeBasisRef:='',DriftBoundPpm:=0,DriftEvidence:='',HistoryBasisRef:='',HistoryUtcLowerMs:=0,
        RequestSubmitted:=FALSE,ResponseReady:=FALSE,HeartbeatSubmitted:=FALSE,ConfigGetSubmitted:=FALSE);
    Checks[22]:=NOT LogicalClock.TimeValid AND LogicalClock.EnqueueAllowed AND NOT LogicalClock.RequestWanted;
    LogicalClock(Reset:=TRUE,PlatformMode:=TRUE,Connected:=TRUE,SessionId:='bad-drift',NowMs:=Tick,SystemUtcMs:=SystemDate,
        TimeBasisRef:='site-hub-1',DriftBoundPpm:=50,DriftEvidence:='',HistoryBasisRef:='',HistoryUtcLowerMs:=0);
    Checks[23]:=(LogicalClock.State=6) AND NOT LogicalClock.EnqueueAllowed;
    LogicalClock(Reset:=TRUE,PlatformMode:=TRUE,Connected:=TRUE,SessionId:='bad-basis',NowMs:=Tick,SystemUtcMs:=SystemDate,
        TimeBasisRef:='site-hub-1',DriftBoundPpm:=50,DriftEvidence:='TEST_FIXTURE_ONLY',HistoryBasisRef:='other-hub',HistoryUtcLowerMs:=1);
    Checks[24]:=(LogicalClock.State=6) AND NOT LogicalClock.EnqueueAllowed;
21: Checks[25]:=LogicalClock.TimeValid;
22: Checks[26]:=NOT LogicalClock.TimeValid AND (LogicalClock.State=4);
23: Checks[27]:=LogicalClock.RequestWanted;
29:
    Checks[28]:=LogicalClock.TimeValid;
    Checks[29]:=LogicalClock.State=2;
    Checks[30]:=LogicalClock.UtcMs>=SavedOutput;
    Checks[31]:=NOT LogicalClock.SendAllowed;
31: Checks[32]:=LogicalClock.SendAllowed;
38:
    Checks[33]:=LogicalClock.TimeValid AND (LogicalClock.UtcMs>=SavedOutput);
    Checks[34]:=(LogicalClock.State=2) AND (LogicalClock.UncertaintyMs<5000);
45: Checks[35]:=(LogicalClock.State=5) AND NOT LogicalClock.TimeValid;
46: Checks[36]:=LogicalClock.RequestWanted AND NOT LogicalClock.TimeValid;
52: Checks[37]:=(LogicalClock.State=4) AND NOT LogicalClock.TimeValid;
53: Checks[38]:=LogicalClock.RequestWanted;
59: Checks[39]:=LogicalClock.TimeValid AND (LogicalClock.UtcMs>=SavedOutput);
61:
    Checks[40]:=LogicalClock.TimeValid AND LogicalClock.SendAllowed AND (LogicalClock.State=2);
    Passed:=0; FailedChecks:=0;
    FOR i:=1 TO 40 DO IF Checks[i] THEN Passed:=Passed+1; ELSE FailedChecks:=FailedChecks+1; END_IF; END_FOR;
    ClockDone:=TRUE;
END_CASE;
Stage:=Stage+1;

END_FUNCTION_BLOCK

(* ---- NG_PollSlot.st ---- *)
FUNCTION_BLOCK NG_PollSlot
VAR_INPUT
    NowMs : ULINT;
    PeriodMs : UDINT;
END_VAR
VAR_OUTPUT
    NominalDueMs : ULINT;
END_VAR
VAR_IN_OUT
    Cursor : NG_SourceCursor;
    Buffer : NG_Buffer;
END_VAR
VAR
    skipped : ULINT;
END_VAR

(* Caller has checked NowMs>=NextDue; O is activation, never completion/UTC. *)
NominalDueMs:=Cursor.NextDueMonoMs;
IF (PeriodMs=0) OR (NowMs<Cursor.NextDueMonoMs) OR (NowMs>ULINT#9007199254740991) THEN Buffer.CaptureStopped:=TRUE; RETURN; END_IF;
skipped:=(NowMs-Cursor.NextDueMonoMs)/TO_ULINT(PeriodMs);
IF skipped>ULINT#9007199254740991-Buffer.MissedPollCyclesTotal THEN Buffer.CounterOverflow:=TRUE; END_IF;
Buffer.MissedPollCyclesTotal:=NG_SafeAdd(Buffer.MissedPollCyclesTotal,skipped);
NominalDueMs:=Cursor.NextDueMonoMs+skipped*TO_ULINT(PeriodMs);
IF NominalDueMs>ULINT#9007199254740991-TO_ULINT(PeriodMs) THEN Buffer.CaptureStopped:=TRUE;
ELSE Cursor.NextDueMonoMs:=NominalDueMs+TO_ULINT(PeriodMs); END_IF;
END_FUNCTION_BLOCK

(* ---- NG_PruneTerminal.st ---- *)
FUNCTION_BLOCK NG_PruneTerminal
VAR_INPUT
    Index : UINT;
END_VAR
VAR_IN_OUT
    Buffer : NG_Buffer;
END_VAR
VAR
    Free : NG_FreeRecord;
    j : UINT;
    r : UINT;
    offset : UINT;
END_VAR
IF (Index=0) OR (Index>64) THEN RETURN; END_IF;
IF Buffer.TerminalOwners[Index].Count=0 THEN RETURN; END_IF;
offset:=(Index-1)*64;
FOR j:=1 TO Buffer.TerminalOwners[Index].Count DO
    r:=Buffer.TerminalRefs[offset+j];
    IF r=0 THEN Buffer.CaptureStopped:=TRUE; Buffer.AccountingComplete:=FALSE; RETURN; END_IF;
    IF (Buffer.RecordGenerations[r]<>Buffer.TerminalRefGenerations[offset+j]) OR (Buffer.RecordStates[r]=0) THEN
        Buffer.CaptureStopped:=TRUE; Buffer.AccountingComplete:=FALSE; RETURN;
    END_IF;
END_FOR;
FOR j:=1 TO Buffer.TerminalOwners[Index].Count DO
    r:=Buffer.TerminalRefs[offset+j];
    IF (r<>0) AND (Buffer.RecordGenerations[r]=Buffer.TerminalRefGenerations[offset+j]) THEN Free(Index:=r,Buffer:=Buffer);
    ELSE Buffer.CaptureStopped:=TRUE; END_IF;
    Buffer.TerminalRefs[offset+j]:=0;
END_FOR;
Buffer.TerminalOwners[Index].Count:=0; Buffer.TerminalOwners[Index].MessageId:='';
Buffer.TombstonePrunedBatchesTotal:=NG_SafeAdd(Buffer.TombstonePrunedBatchesTotal,ULINT#1);
Buffer.DetailTruncated:=TRUE;
END_FUNCTION_BLOCK
